   VAR 
      switching_on_inhibited : Bool := FALSE;
      ready_for_switching_on : Bool := FALSE;
      switched_on : Bool := FALSE;
      operation : Bool := FALSE;
      ars_statusword : Word;
      ars_controlword : Word;
      start_pos : Bool := FALSE;
      start_pos_old : Bool := FALSE;   // ***********************************************************************************************************************Anweisungsteil
      start_pos_man : Bool;
      start_pos_man_old : Bool;
      Fahrauftrag_OK : Bool;
      AFAG_Ist_Wert_in_Grad : Real;
      AFAG_soll_Wert_in_Grad : Real;
      AFAG_soll_Speed_in_Prozent : Int;
      AFAG_soll_Beschleunigung_in_Grad_s : Int;
      abs_rel : Bool;
      R_TRIG_Instance {InstructionName := 'R_TRIG'; LibVersion := '1.0'} : R_TRIG;
      R_TRIG_Q_Tipp_neg : Bool;
      R_TRIG_Instance_1 {InstructionName := 'R_TRIG'; LibVersion := '1.0'} : R_TRIG;
      R_TRIG_Instance_2 {InstructionName := 'R_TRIG'; LibVersion := '1.0'} : R_TRIG;
      TP_Time_Pos_0 {InstructionName := 'TP_TIME'; LibVersion := '1.0'} : TP_TIME;
      TP_Time_Pos_1 {InstructionName := 'TP_TIME'; LibVersion := '1.0'} : TP_TIME;
      TP_Time_Pos_2 {InstructionName := 'TP_TIME'; LibVersion := '1.0'} : TP_TIME;
      TP_Time_Pos_3 {InstructionName := 'TP_TIME'; LibVersion := '1.0'} : TP_TIME;
      TP_Time_Pos_4 {InstructionName := 'TP_TIME'; LibVersion := '1.0'} : TP_TIME;
      TP_Time_Pos_5 {InstructionName := 'TP_TIME'; LibVersion := '1.0'} : TP_TIME;
      TP_Time_Pos_6 {InstructionName := 'TP_TIME'; LibVersion := '1.0'} : TP_TIME;
      TP_Time_Pos_7 {InstructionName := 'TP_TIME'; LibVersion := '1.0'} : TP_TIME;
      TP_Time_Pos_8 {InstructionName := 'TP_TIME'; LibVersion := '1.0'} : TP_TIME;
      TP_Time_Pos_9 {InstructionName := 'TP_TIME'; LibVersion := '1.0'} : TP_TIME;
      TP_Time_Pos_10 {InstructionName := 'TP_TIME'; LibVersion := '1.0'} : TP_TIME;
      TP_Time_Pos_11 {InstructionName := 'TP_TIME'; LibVersion := '1.0'} : TP_TIME;
      TP_Time_Pos_12 {InstructionName := 'TP_TIME'; LibVersion := '1.0'} : TP_TIME;
      TP_Time_Pos_13 {InstructionName := 'TP_TIME'; LibVersion := '1.0'} : TP_TIME;
      TP_Time_Pos_14 {InstructionName := 'TP_TIME'; LibVersion := '1.0'} : TP_TIME;
      TP_Time_Pos_15 {InstructionName := 'TP_TIME'; LibVersion := '1.0'} : TP_TIME;
   END_VAR


BEGIN
	
	
	//Ausgänge zuweisen
	#A_UDT_Afag_soll_Werte.Telegrammkennung := 16#e0;
	#A_Afag_ist_wert_Grad := #AFAG_Ist_Wert_in_Grad;
	#AFAG_Ist_Wert_in_Grad := (DINT_TO_REAL(#E_UDT_Afag_ist_Werte.actual_position)); // / 1.000000e+003;
	#A_UDT_Afag_soll_Werte.Zielposition := REAL_TO_DINT(#AFAG_soll_Wert_in_Grad); // * 1.000000e+003);
	#A_UDT_Afag_soll_Werte.Fahrgeschwindigkeit := INT_TO_DINT(#AFAG_soll_Speed_in_Prozent * (#E_I_Max_Speed_Grad_s / 100));
	#A_UDT_Afag_soll_Werte.Beschleunigung := INT_TO_DINT(#AFAG_soll_Beschleunigung_in_Grad_s);
	#E_A_UDT_Afag_Positionen.A_Softw_ES_min_Grad := 0;
	#E_A_UDT_Afag_Positionen.A_Softw_ES_max_Grad := 360000;
	#E_A_UDT_Afag_Positionen.A_Max_Speed_Grad_s := #E_I_Max_Speed_Grad_s;
	#E_A_UDT_Afag_Positionen.A_Max_Beschleunigung_Grad_s := #E_I_Max_Beschleunigung_Grad_s;
	
	
	//************************************************************************************************
	
	//Lesen Statusword
	//Einlesen des Istzustands der Statemachine
	
	//    #DB_nr_actual_value_word:= INT_TO_WORD(#DB_nr_actual_value);
	//    #ars_statusword := PEEK_WORD (area := 16#84,
	//                                  dbNumber :=#DB_nr_actual_value_word,
	//                                  byteOffset := 2);
	#ars_statusword := #E_UDT_Afag_ist_Werte.PROFIDRIVE_Statusword;
	
	//Lesen Controlword
	//
	//  #DB_nr_position_word:=  INT_TO_WORD(#DB_nr_position);
	//  #ars_controlword := PEEK_WORD (area := 16#84,
	//                                  dbNumber :=#DB_nr_position_word,
	//                                  byteOffset := 2);
	
	// #ars_controlword := #A_UDT_Afag_soll_Werte.PROFIDRIVE_Controlword;
	
	//Steuern der Statemachine, S1 -> S2 -> S3 -> S4
	
	IF (#switching_on_inhibited                          //wenn state "switching_on_inhibited"
	    AND #E_drive_enable)                             //und  Reglerfreigabe
	THEN
	    #ars_controlword := 16#0406;              //dann state "ready_for_switching_on" anfordern,
	ELSIF (#switching_on_inhibited                     //
	    AND (NOT (#E_drive_enable)))                      //wenn Reglerfreigabe aus,
	THEN
	    #ars_controlword := 16#0400;              //dann state "switching_on_inhibited" anfordern.
	END_IF;
	
	IF (#ready_for_switching_on                          //wenn state "ready_for_switching_on"
	    AND #E_drive_enable)                             //und Reglerfeigabe
	THEN
	    #ars_controlword := 16#0407;              //dann state "switched_on" anfordern,
	ELSIF (#ready_for_switching_on                     //
	    AND (NOT (#E_drive_enable)))                      //wenn Reglerfeigabe aus,
	THEN
	    #ars_controlword := 16#0400;              //dann state "switching_on_inhibited" anfordern.
	END_IF;
	
	IF (#switched_on                                     //wenn state "switched_on"
	    AND #E_drive_enable)                             //und Reglerfeigabe
	THEN
	    #ars_controlword := 16#040f;              //dann state "operation" anfordern,
	ELSIF (#switched_on                                //
	    AND (NOT (#E_drive_enable)))                      //wenn Reglerfeigabe aus,
	THEN
	    #ars_controlword := 16#0400;              //dann state "switching_on_inhibited" anfordern.
	END_IF;
	
	IF (#operation                                       //wenn state "operation"
	    AND (NOT (#E_drive_enable)))                      //und keine Reglerfeigabe
	THEN
	    #ars_controlword := 16#040e;              //dann state "switching_on_inhibited" anfordern.
	END_IF;
	
	//************************************************************************************************
	
	//Kommandos über digitale Eingänge
	// Bit 10 (control by plc) im Controlword muss immer gesetzt sein
	
	IF #E_start_homing
	THEN
	    #ars_controlword := (#ars_controlword OR 16#0C00);    //Setzen Bit 11 im STW1
	ELSE
	    #ars_controlword := (#ars_controlword & 16#f7ff);
	END_IF;
	
	IF (#Fahrauftrag_OK = 1) THEN
	    IF (#start_pos_old <> #start_pos) OR (#start_pos_man_old <> #start_pos_man)
	    THEN
	        IF #start_pos OR #start_pos_man
	        THEN
	            #ars_controlword := (#ars_controlword OR 16#0440);    //Setzen Bit 6 im STW1
	        ELSE
	            #ars_controlword := (#ars_controlword & 16#ffbf);
	        END_IF;
	    END_IF;
	    
	    #start_pos_old := #start_pos;
	    #start_pos_man_old := #start_pos_man;
	    
	END_IF;
	
	
	
	
	IF #abs_rel
	THEN
	    #ars_controlword := (#ars_controlword OR 16#1400);   //Setzen Bit 12 im STW1
	ELSE
	    #ars_controlword := (#ars_controlword & 16#efff);
	END_IF;
	
	IF #E_change_immediatly
	THEN
	    #ars_controlword := (#ars_controlword OR 16#2400);   //Setzen Bit 13 im STW1
	ELSE
	    #ars_controlword := (#ars_controlword & 16#dfff);
	END_IF;
	
	IF #E_intermediate_stop
	THEN
	    #ars_controlword := (#ars_controlword & 16#ffdf);   //Rücksetzen Bit 5 im STW1
	ELSE
	    #ars_controlword := (#ars_controlword OR 16#0420);
	END_IF;
	
	IF #E_hold
	THEN
	    #ars_controlword := (#ars_controlword & 16#ffef);    //Rücksetzen Bit 4 im STW1
	    #ars_controlword := (#ars_controlword & 16#feff);    //Rücksetzen jog_pos
	    #ars_controlword := (#ars_controlword & 16#fdff);    //Rücksetzen jog_neg
	ELSE
	    #ars_controlword := (#ars_controlword OR 16#0410);
	END_IF;
	
	IF (#E_jog_pos AND NOT #E_hold)
	THEN
	    #ars_controlword := (#ars_controlword OR 16#0500);    //Setzen Bit 8 im STW1
	ELSE
	    #ars_controlword := (#ars_controlword & 16#feff);
	END_IF;
	
	IF (#E_jog_neg AND NOT #E_hold)
	THEN
	    #ars_controlword := (#ars_controlword OR 16#0600);    //Setzen Bit 9 im STW1
	ELSE
	    #ars_controlword := (#ars_controlword & 16#fdff);
	END_IF;
	
	IF #E_fault_reset
	THEN
	    #ars_controlword := (#ars_controlword OR 16#0480);    //Setzen Bit 7 im STW1
	ELSE
	    #ars_controlword := (#ars_controlword & 16#ff7f);
	END_IF;
	
	
	//************************************************************************************************
	
	//Setzen digitaler Ausgänge
	
	IF #operation
	THEN
	    #A_drive_enable_ok := TRUE;
	ELSE
	    #A_drive_enable_ok := FALSE;
	END_IF;
	
	IF ((#ars_statusword & 16#0800) = 16#0800)    //Bit 11 vom ZSW1
	THEN
	    #A_home_valid := TRUE;
	ELSE
	    #A_home_valid := FALSE;
	END_IF;
	
	IF ((#ars_statusword & 16#0400) = 16#0400)    //Bit 10 vom ZSW1
	THEN
	    #A_pos_ok := TRUE;
	ELSE
	    #A_pos_ok := FALSE;
	END_IF;
	
	IF ((#ars_statusword & 16#2000) = 16#2000)    //Bit 13 vom ZSW1
	THEN
	    #A_velo_zero := TRUE;
	ELSE
	    #A_velo_zero := FALSE;
	END_IF;
	
	IF ((#ars_statusword & 16#0008) = 16#0008)    //Bit 3 vom ZSW1
	THEN
	    #A_fault := TRUE;
	ELSE
	    #A_fault := FALSE;
	END_IF;
	
	//************************************************************************************************
	
	//Schreiben Controlword
	
	//  POKE (area := 16#84,
	//        dbNumber := #DB_nr_position_word,
	//        byteOffset := 2,
	//        value := #ars_controlword );
	
	#A_UDT_Afag_soll_Werte.PROFIDRIVE_Controlword := #ars_controlword;
	
	
	// Achse mit Position Starten
	// Position[0]
	
	    IF #E_A_UDT_Afag_Positionen.Start_POS_Position[0] THEN
	    #AFAG_soll_Wert_in_Grad := #E_A_UDT_Afag_Positionen.Soll_Wert_in_Grad_Position[0];
	    #AFAG_soll_Beschleunigung_in_Grad_s := #E_A_UDT_Afag_Positionen.Soll_Beschleunigung_in_Grad_s_Position[0];
	    #start_pos := true;
	    
	    #AFAG_soll_Speed_in_Prozent := #E_A_UDT_Afag_Positionen.Soll_Speed_in_Prozent_Position[0];
	END_IF;
	
	// Position[1]
	
	IF #E_A_UDT_Afag_Positionen.Start_POS_Position[1] THEN
	    #AFAG_soll_Wert_in_Grad := #E_A_UDT_Afag_Positionen.Soll_Wert_in_Grad_Position[1];
	    #AFAG_soll_Beschleunigung_in_Grad_s := #E_A_UDT_Afag_Positionen.Soll_Beschleunigung_in_Grad_s_Position[1];
	    #start_pos := true;
	    
	    #AFAG_soll_Speed_in_Prozent := #E_A_UDT_Afag_Positionen.Soll_Speed_in_Prozent_Position[1];
	END_IF;
	
	
	// Position 2
	
	IF #E_A_UDT_Afag_Positionen.Start_POS_Position[2] THEN
	    #AFAG_soll_Wert_in_Grad := #E_A_UDT_Afag_Positionen.Soll_Wert_in_Grad_Position[2];
	    #AFAG_soll_Beschleunigung_in_Grad_s := #E_A_UDT_Afag_Positionen.Soll_Beschleunigung_in_Grad_s_Position[2];
	    #start_pos := true;
	    
	    #AFAG_soll_Speed_in_Prozent := #E_A_UDT_Afag_Positionen.Soll_Speed_in_Prozent_Position[2];
	END_IF;
	
	// Position 3
	
	IF #E_A_UDT_Afag_Positionen.Start_POS_Position[3] THEN
	    #AFAG_soll_Wert_in_Grad := #E_A_UDT_Afag_Positionen.Soll_Wert_in_Grad_Position[3];
	    #AFAG_soll_Beschleunigung_in_Grad_s := #E_A_UDT_Afag_Positionen.Soll_Beschleunigung_in_Grad_s_Position[3];
	    #start_pos := true;
	    
	    #AFAG_soll_Speed_in_Prozent := #E_A_UDT_Afag_Positionen.Soll_Speed_in_Prozent_Position[3];
	END_IF;
	
	// Position 4
	
	IF #E_A_UDT_Afag_Positionen.Start_POS_Position[4] THEN
	    #AFAG_soll_Wert_in_Grad := #E_A_UDT_Afag_Positionen.Soll_Wert_in_Grad_Position[4];
	    #AFAG_soll_Beschleunigung_in_Grad_s := #E_A_UDT_Afag_Positionen.Soll_Beschleunigung_in_Grad_s_Position[4];
	    #start_pos := true;
	    
	    #AFAG_soll_Speed_in_Prozent := #E_A_UDT_Afag_Positionen.Soll_Speed_in_Prozent_Position[4];
	END_IF;
	
	// Position 5
	
	IF #E_A_UDT_Afag_Positionen.Start_POS_Position[5] THEN
	    #AFAG_soll_Wert_in_Grad := #E_A_UDT_Afag_Positionen.Soll_Wert_in_Grad_Position[5];
	    #AFAG_soll_Beschleunigung_in_Grad_s := #E_A_UDT_Afag_Positionen.Soll_Beschleunigung_in_Grad_s_Position[5];
	    #start_pos := true;
	    
	    #AFAG_soll_Speed_in_Prozent := #E_A_UDT_Afag_Positionen.Soll_Speed_in_Prozent_Position[5];
	END_IF;
	
	// Position 6
	
	IF #E_A_UDT_Afag_Positionen.Start_POS_Position[6] THEN
	    #AFAG_soll_Wert_in_Grad := #E_A_UDT_Afag_Positionen.Soll_Wert_in_Grad_Position[6];
	    #AFAG_soll_Beschleunigung_in_Grad_s := #E_A_UDT_Afag_Positionen.Soll_Beschleunigung_in_Grad_s_Position[6];
	    #start_pos := true;
	    
	    #AFAG_soll_Speed_in_Prozent := #E_A_UDT_Afag_Positionen.Soll_Speed_in_Prozent_Position[6];
	END_IF;
	
	// Position 7
	
	IF #E_A_UDT_Afag_Positionen.Start_POS_Position[7] THEN
	    #AFAG_soll_Wert_in_Grad := #E_A_UDT_Afag_Positionen.Soll_Wert_in_Grad_Position[7];
	    #AFAG_soll_Beschleunigung_in_Grad_s := #E_A_UDT_Afag_Positionen.Soll_Beschleunigung_in_Grad_s_Position[7];
	    #start_pos := true;
	    
	    #AFAG_soll_Speed_in_Prozent := #E_A_UDT_Afag_Positionen.Soll_Speed_in_Prozent_Position[7];
	END_IF;
	
	// Position 8
	
	IF #E_A_UDT_Afag_Positionen.Start_POS_Position[8] THEN
	    #AFAG_soll_Wert_in_Grad := #E_A_UDT_Afag_Positionen.Soll_Wert_in_Grad_Position[8];
	    #AFAG_soll_Beschleunigung_in_Grad_s := #E_A_UDT_Afag_Positionen.Soll_Beschleunigung_in_Grad_s_Position[8];
	    #start_pos := true;
	    
	    #AFAG_soll_Speed_in_Prozent := #E_A_UDT_Afag_Positionen.Soll_Speed_in_Prozent_Position[8];
	END_IF;
	
	// Position 9
	
	IF #E_A_UDT_Afag_Positionen.Start_POS_Position[9] THEN
	    #AFAG_soll_Wert_in_Grad := #E_A_UDT_Afag_Positionen.Soll_Wert_in_Grad_Position[9];
	    #AFAG_soll_Beschleunigung_in_Grad_s := #E_A_UDT_Afag_Positionen.Soll_Beschleunigung_in_Grad_s_Position[9];
	    #start_pos := true;
	   
	    #AFAG_soll_Speed_in_Prozent := #E_A_UDT_Afag_Positionen.Soll_Speed_in_Prozent_Position[9];
	END_IF;
	
	// Position 10
	
	IF #E_A_UDT_Afag_Positionen.Start_POS_Position[10] THEN
	    #AFAG_soll_Wert_in_Grad := #E_A_UDT_Afag_Positionen.Soll_Wert_in_Grad_Position[10];
	    #AFAG_soll_Beschleunigung_in_Grad_s := #E_A_UDT_Afag_Positionen.Soll_Beschleunigung_in_Grad_s_Position[10];
	    #start_pos := true;
	    
	    #AFAG_soll_Speed_in_Prozent := #E_A_UDT_Afag_Positionen.Soll_Speed_in_Prozent_Position[10];
	END_IF;
	
	// Position 11
	
	IF #E_A_UDT_Afag_Positionen.Start_POS_Position[11] THEN
	    #AFAG_soll_Wert_in_Grad := #E_A_UDT_Afag_Positionen.Soll_Wert_in_Grad_Position[11];
	    #AFAG_soll_Beschleunigung_in_Grad_s := #E_A_UDT_Afag_Positionen.Soll_Beschleunigung_in_Grad_s_Position[11];
	    #start_pos := true;
	    
	    #AFAG_soll_Speed_in_Prozent := #E_A_UDT_Afag_Positionen.Soll_Speed_in_Prozent_Position[11];
	END_IF;
	
	// Position 12
	
	IF #E_A_UDT_Afag_Positionen.Start_POS_Position[12] THEN
	    #AFAG_soll_Wert_in_Grad := #E_A_UDT_Afag_Positionen.Soll_Wert_in_Grad_Position[12];
	    #AFAG_soll_Beschleunigung_in_Grad_s := #E_A_UDT_Afag_Positionen.Soll_Beschleunigung_in_Grad_s_Position[12];
	    #start_pos := true;
	    
	    #AFAG_soll_Speed_in_Prozent := #E_A_UDT_Afag_Positionen.Soll_Speed_in_Prozent_Position[12];
	END_IF;
	
	// Position 13
	
	IF #E_A_UDT_Afag_Positionen.Start_POS_Position[13] THEN
	    #AFAG_soll_Wert_in_Grad := #E_A_UDT_Afag_Positionen.Soll_Wert_in_Grad_Position[13];
	    #AFAG_soll_Beschleunigung_in_Grad_s := #E_A_UDT_Afag_Positionen.Soll_Beschleunigung_in_Grad_s_Position[13];
	    #start_pos := true;
	    
	    #AFAG_soll_Speed_in_Prozent := #E_A_UDT_Afag_Positionen.Soll_Speed_in_Prozent_Position[13];
	END_IF;
	
	// Position 14
	
	IF #E_A_UDT_Afag_Positionen.Start_POS_Position[14] THEN
	    #AFAG_soll_Wert_in_Grad := #E_A_UDT_Afag_Positionen.Soll_Wert_in_Grad_Position[14];
	    #AFAG_soll_Beschleunigung_in_Grad_s := #E_A_UDT_Afag_Positionen.Soll_Beschleunigung_in_Grad_s_Position[14];
	    #start_pos := true;
	    
	    #AFAG_soll_Speed_in_Prozent := #E_A_UDT_Afag_Positionen.Soll_Speed_in_Prozent_Position[14];
	END_IF;
	
	// Position 15
	
	IF #E_A_UDT_Afag_Positionen.Start_POS_Position[15] THEN
	    #AFAG_soll_Wert_in_Grad := #E_A_UDT_Afag_Positionen.Soll_Wert_in_Grad_Position[15];
	    #AFAG_soll_Beschleunigung_in_Grad_s := #E_A_UDT_Afag_Positionen.Soll_Beschleunigung_in_Grad_s_Position[15];
	    #start_pos := true;
	    
	    #AFAG_soll_Speed_in_Prozent := #E_A_UDT_Afag_Positionen.Soll_Speed_in_Prozent_Position[15];
	END_IF;
	
	// Manuelle Geschwindigkeitsanpassung
	IF #E_BA_Manuell = TRUE THEN
	   #AFAG_soll_Speed_in_Prozent := #E_I_Manuell_Geschwindigkeit_Prozent;
	   #AFAG_soll_Beschleunigung_in_Grad_s := 1000;
	END_IF;
	
	IF( (#E_A_UDT_Afag_Positionen.Start_POS_Position[0] AND #E_A_UDT_Afag_Positionen.POS_OK_Position[0])OR
	   (#E_A_UDT_Afag_Positionen.Start_POS_Position[1]AND #E_A_UDT_Afag_Positionen.POS_OK_Position[1])OR
	   (#E_A_UDT_Afag_Positionen.Start_POS_Position[2]AND #E_A_UDT_Afag_Positionen.POS_OK_Position[2])OR
	   (#E_A_UDT_Afag_Positionen.Start_POS_Position[3]AND #E_A_UDT_Afag_Positionen.POS_OK_Position[3])OR
	   (#E_A_UDT_Afag_Positionen.Start_POS_Position[4]AND #E_A_UDT_Afag_Positionen.POS_OK_Position[4])OR
	   (#E_A_UDT_Afag_Positionen.Start_POS_Position[5]AND #E_A_UDT_Afag_Positionen.POS_OK_Position[5])OR
	   (#E_A_UDT_Afag_Positionen.Start_POS_Position[6]AND #E_A_UDT_Afag_Positionen.POS_OK_Position[6])OR
	   (#E_A_UDT_Afag_Positionen.Start_POS_Position[7]AND #E_A_UDT_Afag_Positionen.POS_OK_Position[7])OR
	   (#E_A_UDT_Afag_Positionen.Start_POS_Position[8]AND #E_A_UDT_Afag_Positionen.POS_OK_Position[8])OR
	   (#E_A_UDT_Afag_Positionen.Start_POS_Position[9]AND #E_A_UDT_Afag_Positionen.POS_OK_Position[9])OR
	   (#E_A_UDT_Afag_Positionen.Start_POS_Position[10]AND #E_A_UDT_Afag_Positionen.POS_OK_Position[10])OR
	   (#E_A_UDT_Afag_Positionen.Start_POS_Position[11]AND #E_A_UDT_Afag_Positionen.POS_OK_Position[11])OR
	   (#E_A_UDT_Afag_Positionen.Start_POS_Position[12]AND #E_A_UDT_Afag_Positionen.POS_OK_Position[12])OR
	   (#E_A_UDT_Afag_Positionen.Start_POS_Position[13]AND #E_A_UDT_Afag_Positionen.POS_OK_Position[13])OR
	   (#E_A_UDT_Afag_Positionen.Start_POS_Position[14]AND #E_A_UDT_Afag_Positionen.POS_OK_Position[14])OR
	   (#E_A_UDT_Afag_Positionen.Start_POS_Position[15]AND #E_A_UDT_Afag_Positionen.POS_OK_Position[15])OR
	    #E_Richten_reset_FRG)
	THEN
	    #start_pos := 0;
	    #E_A_UDT_Afag_Positionen.Start_POS_Position[0] := 0;
	    #E_A_UDT_Afag_Positionen.Start_POS_Position[1] := 0;
	    #E_A_UDT_Afag_Positionen.Start_POS_Position[2] := 0;
	    #E_A_UDT_Afag_Positionen.Start_POS_Position[3] := 0;
	    #E_A_UDT_Afag_Positionen.Start_POS_Position[4] := 0;
	    #E_A_UDT_Afag_Positionen.Start_POS_Position[5] := 0;
	    #E_A_UDT_Afag_Positionen.Start_POS_Position[6] := 0;
	    #E_A_UDT_Afag_Positionen.Start_POS_Position[7] := 0;
	    #E_A_UDT_Afag_Positionen.Start_POS_Position[8] := 0;
	    #E_A_UDT_Afag_Positionen.Start_POS_Position[9] := 0;
	    #E_A_UDT_Afag_Positionen.Start_POS_Position[10] := 0;
	    #E_A_UDT_Afag_Positionen.Start_POS_Position[11] := 0;
	    #E_A_UDT_Afag_Positionen.Start_POS_Position[12] := 0;
	    #E_A_UDT_Afag_Positionen.Start_POS_Position[13] := 0;
	    #E_A_UDT_Afag_Positionen.Start_POS_Position[14] := 0;
	    #E_A_UDT_Afag_Positionen.Start_POS_Position[15] := 0;
	    #E_A_UDT_Afag_Positionen.POS_OK_Position[15] := 0;
	END_IF;
	
	
	// Achse Positionsrückmeldung
	
	IF #E_A_UDT_Afag_Positionen.Start_POS_Position[0] AND #A_pos_ok
	THEN
	    #E_A_UDT_Afag_Positionen.POS_OK_Position[0] := 1;
	ELSE
	    #E_A_UDT_Afag_Positionen.POS_OK_Position[0] := 0;
	END_IF;
	
	IF #E_A_UDT_Afag_Positionen.Start_POS_Position[1] AND #A_pos_ok
	THEN
	    #E_A_UDT_Afag_Positionen.POS_OK_Position[1] := 1;
	ELSE
	    #E_A_UDT_Afag_Positionen.POS_OK_Position[1] := 0;
	END_IF;
	
	IF #E_A_UDT_Afag_Positionen.Start_POS_Position[2] AND #A_pos_ok
	THEN
	    #E_A_UDT_Afag_Positionen.POS_OK_Position[2] := 1;
	ELSE
	    #E_A_UDT_Afag_Positionen.POS_OK_Position[2] := 0;
	END_IF;
	
	IF #E_A_UDT_Afag_Positionen.Start_POS_Position[3] AND #A_pos_ok
	THEN
	    #E_A_UDT_Afag_Positionen.POS_OK_Position[3] := 1;
	ELSE
	    #E_A_UDT_Afag_Positionen.POS_OK_Position[3] := 0;
	END_IF;
	
	IF #E_A_UDT_Afag_Positionen.Start_POS_Position[4] AND #A_pos_ok
	THEN
	    #E_A_UDT_Afag_Positionen.POS_OK_Position[4] := 1;
	ELSE
	    #E_A_UDT_Afag_Positionen.POS_OK_Position[4] := 0;
	END_IF;
	
	IF #E_A_UDT_Afag_Positionen.Start_POS_Position[5] AND #A_pos_ok
	THEN
	    #E_A_UDT_Afag_Positionen.POS_OK_Position[5] := 1;
	ELSE
	    #E_A_UDT_Afag_Positionen.POS_OK_Position[5] := 0;
	END_IF;
	
	IF #E_A_UDT_Afag_Positionen.Start_POS_Position[6] AND #A_pos_ok
	THEN
	    #E_A_UDT_Afag_Positionen.POS_OK_Position[6] := 1;
	ELSE
	    #E_A_UDT_Afag_Positionen.POS_OK_Position[6] := 0;
	END_IF;
	
	IF #E_A_UDT_Afag_Positionen.Start_POS_Position[7] AND #A_pos_ok
	THEN
	    #E_A_UDT_Afag_Positionen.POS_OK_Position[7] := 1;
	ELSE
	    #E_A_UDT_Afag_Positionen.POS_OK_Position[7] := 0;
	END_IF;
	
	IF #E_A_UDT_Afag_Positionen.Start_POS_Position[8] AND #A_pos_ok
	THEN
	    #E_A_UDT_Afag_Positionen.POS_OK_Position[8] := 1;
	ELSE
	    #E_A_UDT_Afag_Positionen.POS_OK_Position[8] := 0;
	END_IF;
	
	IF #E_A_UDT_Afag_Positionen.Start_POS_Position[9] AND #A_pos_ok
	THEN
	    #E_A_UDT_Afag_Positionen.POS_OK_Position[9] := 1;
	ELSE
	    #E_A_UDT_Afag_Positionen.POS_OK_Position[9] := 0;
	END_IF;
	
	IF #E_A_UDT_Afag_Positionen.Start_POS_Position[10] AND #A_pos_ok
	THEN
	    #E_A_UDT_Afag_Positionen.POS_OK_Position[10] := 1;
	ELSE
	    #E_A_UDT_Afag_Positionen.POS_OK_Position[10] := 0;
	END_IF;
	
	IF #E_A_UDT_Afag_Positionen.Start_POS_Position[11] AND #A_pos_ok
	THEN
	    #E_A_UDT_Afag_Positionen.POS_OK_Position[11] := 1;
	ELSE
	    #E_A_UDT_Afag_Positionen.POS_OK_Position[11] := 0;
	END_IF;
	
	IF #E_A_UDT_Afag_Positionen.Start_POS_Position[12] AND #A_pos_ok
	THEN
	    #E_A_UDT_Afag_Positionen.POS_OK_Position[12] := 1;
	ELSE
	    #E_A_UDT_Afag_Positionen.POS_OK_Position[12] := 0;
	END_IF;
	
	IF #E_A_UDT_Afag_Positionen.Start_POS_Position[13] AND #A_pos_ok
	THEN
	    #E_A_UDT_Afag_Positionen.POS_OK_Position[13] := 1;
	ELSE
	    #E_A_UDT_Afag_Positionen.POS_OK_Position[13] := 0;
	END_IF;
	
	IF #E_A_UDT_Afag_Positionen.Start_POS_Position[14] AND #A_pos_ok
	THEN
	    #E_A_UDT_Afag_Positionen.POS_OK_Position[14] := 1;
	ELSE
	    #E_A_UDT_Afag_Positionen.POS_OK_Position[14] := 0;
	END_IF;
	
	IF #E_A_UDT_Afag_Positionen.Start_POS_Position[15] AND #A_pos_ok
	THEN
	    #E_A_UDT_Afag_Positionen.POS_OK_Position[15] := 1;
	ELSE
	    #E_A_UDT_Afag_Positionen.POS_OK_Position[15] := 0;
	END_IF;
	
	IF
	    (#E_A_UDT_Afag_Positionen.Start_POS_Position[0]) OR
	    (#E_A_UDT_Afag_Positionen.Start_POS_Position[1]) OR
	    (#E_A_UDT_Afag_Positionen.Start_POS_Position[2]) OR
	    (#E_A_UDT_Afag_Positionen.Start_POS_Position[3]) OR
	    (#E_A_UDT_Afag_Positionen.Start_POS_Position[4]) OR
	    (#E_A_UDT_Afag_Positionen.Start_POS_Position[5]) OR
	    (#E_A_UDT_Afag_Positionen.Start_POS_Position[6]) OR
	    (#E_A_UDT_Afag_Positionen.Start_POS_Position[7]) OR
	    (#E_A_UDT_Afag_Positionen.Start_POS_Position[8]) OR
	    (#E_A_UDT_Afag_Positionen.Start_POS_Position[9]) OR
	    (#E_A_UDT_Afag_Positionen.Start_POS_Position[10]) OR
	    (#E_A_UDT_Afag_Positionen.Start_POS_Position[11]) OR
	    (#E_A_UDT_Afag_Positionen.Start_POS_Position[12]) OR
	    (#E_A_UDT_Afag_Positionen.Start_POS_Position[13]) OR
	    (#E_A_UDT_Afag_Positionen.Start_POS_Position[14]) OR
	    (#E_A_UDT_Afag_Positionen.Start_POS_Position[15]) OR
	    (#start_pos)
	THEN
	    #A_Fahrauftrag_Aktiv := 1;
	ELSE
	    #A_Fahrauftrag_Aktiv := 0;
	END_IF;
	
	
	
	
	//Reset Start pos
	IF ((#A_pos_ok = true) OR (#A_drive_enable_ok = FALSE) OR (#E_fault_reset = TRUE))
	THEN
	    #start_pos_man := false;
	    #abs_rel := true;
	END_IF;
	
	//Tipp pos
	#R_TRIG_Instance(CLK:=#E_Tipp_pos);
	IF (#R_TRIG_Instance.Q AND NOT #start_pos_man)
	THEN
	    #AFAG_soll_Wert_in_Grad := #E_R_Verfahrweg_Grad;
	    #start_pos_man := TRUE;
	END_IF;
	
	//Tipp neg
	#R_TRIG_Instance_1(CLK:=#E_Tipp_neg);
	IF (#R_TRIG_Instance_1.Q AND NOT #start_pos_man)
	THEN
	    #AFAG_soll_Wert_in_Grad := #E_R_Verfahrweg_Grad;
	    #start_pos_man := TRUE;
	END_IF;
	
	//absolut verfahren
	#R_TRIG_Instance_2(CLK:=#E_Start_pos_man);
	IF(#R_TRIG_Instance_2.Q AND NOT #start_pos_man)
	THEN
	    #AFAG_soll_Wert_in_Grad := #E_R_Afag_soll_wert_man_Grad;
	    #start_pos_man := TRUE;
	    #abs_rel := false;
	END_IF;
	
	// keine Endlagenüberwachung bei Drehachse
	// Überwachung Fahrauftrag
	    #Fahrauftrag_OK := TRUE;
	 
	    
	//Einlesen des Istzustands der Statemachine
	   IF ((#ars_statusword & 16#0047) = 16#0040)
	        THEN #switching_on_inhibited := TRUE;
	        ELSE #switching_on_inhibited := FALSE;
	    END_IF;
	
	    IF ((#ars_statusword & 16#0047) = 16#0001)
	        THEN #ready_for_switching_on:= TRUE;
	        ELSE #ready_for_switching_on:= FALSE;
	    END_IF;
	     
	    IF ((#ars_statusword & 16#0047) = 16#0003)
	        THEN #switched_on:= TRUE;
	        ELSE #switched_on:= FALSE;
	    END_IF;
	
	    IF ((#ars_statusword & 16#0047) = 16#0007)
	        THEN #operation:= TRUE;
	        ELSE #operation:= FALSE;
	    END_IF;    
	
	
	
	    
	    
END_FUNCTION_BLOCK

FUNCTION_BLOCK "BB_Ansteuerung_Afag_offen_V02.3"
TITLE = 'FB Positionierbetrieb'
{ S7_Optimized_Access := 'TRUE' }
AUTHOR : Essmann
FAMILY : metronix
NAME : position
VERSION : 1.1
//Der Baustein kann nicht rückübersetzt und unter STEP7 bearbeitet werden.  Der Baustein kann nur als Quelle im Ordner "Quellen" bearbeitet werden.    IO-Variablen  
   VAR_INPUT 
      drive_enable : Bool := FALSE;
      start_homing : Bool := FALSE;
      start_pos : Bool := FALSE;
      abs_rel : Bool := FALSE;
      change_immediatly : Bool := FALSE;
      intermediate_stop : Bool := FALSE;
      hold : Bool := FALSE;
      jog_pos : Bool := FALSE;
      jog_neg : Bool := FALSE;
      fault_reset : Bool := FALSE;
      E_Afag_ist_Werte : "Afag_ist_Werte";
   END_VAR

   VAR_OUTPUT 
      drive_enable_ok : Bool := FALSE;
      home_valid : Bool := FALSE;
      pos_ok : Bool := FALSE;
      velo_zero : Bool := FALSE;
      fault : Bool := FALSE;   // statische Variablen
   END_VAR

   VAR_IN_OUT 
      A_Afag_soll_Werte : "Afag_soll_Werte";
   END_VAR

   VAR 
      DB_nr_position_word : Word;
      DB_nr_actual_value_word : Word;
      switching_on_inhibited : Bool := FALSE;
      ready_for_switching_on : Bool := FALSE;
      switched_on : Bool := FALSE;
      operation : Bool := FALSE;
      ars_statusword : Word;
      ars_controlword : Word;
      start_pos_old : Bool := FALSE;   // ***********************************************************************************************************************Anweisungsteil
   END_VAR


BEGIN
	
	
	//Lesen Statusword
	//Einlesen des Istzustands der Statemachine
	    
	 //    #DB_nr_actual_value_word:= INT_TO_WORD(#DB_nr_actual_value);
	 //    #ars_statusword := PEEK_WORD (area := 16#84,
	 //                                  dbNumber :=#DB_nr_actual_value_word,
	 //                                  byteOffset := 2);
	 
	 #A_Afag_soll_Werte.Telegrammkennung:= 16#e0;
	 
	 
	 #ars_statusword := #E_Afag_ist_Werte.PROFIDRIVE_Statusword;
	
	   IF ((#ars_statusword & 16#0047) = 16#0040)
	        THEN #switching_on_inhibited := TRUE;
	        ELSE #switching_on_inhibited := FALSE;
	    END_IF;
	
	    IF ((#ars_statusword & 16#0047) = 16#0001)
	        THEN #ready_for_switching_on:= TRUE;
	        ELSE #ready_for_switching_on:= FALSE;
	    END_IF;
	     
	    IF ((#ars_statusword & 16#0047) = 16#0003)
	        THEN #switched_on:= TRUE;
	        ELSE #switched_on:= FALSE;
	    END_IF;
	
	    IF ((#ars_statusword & 16#0047) = 16#0007)
	        THEN #operation:= TRUE;
	        ELSE #operation:= FALSE;
	    END_IF;    
	
	
	//************************************************************************************************
	
	//Lesen Controlword
	//
	 //  #DB_nr_position_word:=  INT_TO_WORD(#DB_nr_position);
	 //  #ars_controlword := PEEK_WORD (area := 16#84,
	 //                                  dbNumber :=#DB_nr_position_word,
	 //                                  byteOffset := 2);
	    
	    #ars_controlword := #A_Afag_soll_Werte.PROFIDRIVE_Controlword;
	    
	//Steuern der Statemachine, S1 -> S2 -> S3 -> S4
	
	  IF (#switching_on_inhibited                          //wenn state "switching_on_inhibited"
	        AND #drive_enable)                             //und  Reglerfreigabe
	        THEN #ars_controlword := 16#0406;              //dann state "ready_for_switching_on" anfordern,
	    ELSIF (#switching_on_inhibited                     //
	        AND (NOT(#drive_enable)))                      //wenn Reglerfreigabe aus,
	        THEN #ars_controlword := 16#0400;              //dann state "switching_on_inhibited" anfordern.
	  END_IF;                                             
	
	  IF (#ready_for_switching_on                          //wenn state "ready_for_switching_on"
	        AND #drive_enable)                             //und Reglerfeigabe
	        THEN #ars_controlword := 16#0407;              //dann state "switched_on" anfordern,
	    ELSIF (#ready_for_switching_on                     //
	        AND (NOT(#drive_enable)))                      //wenn Reglerfeigabe aus,
	        THEN #ars_controlword := 16#0400;              //dann state "switching_on_inhibited" anfordern.
	  END_IF;
	
	  IF (#switched_on                                     //wenn state "switched_on"
	        AND #drive_enable)                             //und Reglerfeigabe
	        THEN #ars_controlword := 16#040f;              //dann state "operation" anfordern,
	    ELSIF (#switched_on                                //
	        AND (NOT(#drive_enable)))                      //wenn Reglerfeigabe aus,
	        THEN #ars_controlword := 16#0400;              //dann state "switching_on_inhibited" anfordern.
	  END_IF;
	
	  IF (#operation                                       //wenn state "operation"
	        AND (NOT(#drive_enable)))                      //und keine Reglerfeigabe
	        THEN #ars_controlword := 16#040e;              //dann state "switching_on_inhibited" anfordern.
	  END_IF;
	
	//************************************************************************************************
	
	//Kommandos über digitale Eingänge
	// Bit 10 (control by plc) im Controlword muss immer gesetzt sein
	
	    IF #start_homing
	        THEN #ars_controlword := (#ars_controlword OR 16#0C00);    //Setzen Bit 11 im STW1
	        ELSE #ars_controlword := (#ars_controlword  & 16#f7ff);
	    END_IF;
	
	    IF #start_pos_old <> #start_pos
	        THEN IF #start_pos 
	                 THEN #ars_controlword := (#ars_controlword OR 16#0440);    //Setzen Bit 6 im STW1
	                 ELSE #ars_controlword := (#ars_controlword  & 16#ffbf);
	             END_IF;
	    END_IF;
	
	    #start_pos_old := #start_pos;
	
	    IF #abs_rel
	        THEN #ars_controlword := (#ars_controlword OR 16#1400);   //Setzen Bit 12 im STW1
	        ELSE #ars_controlword := (#ars_controlword  & 16#efff);
	    END_IF;
	    
	    IF #change_immediatly
	        THEN #ars_controlword := (#ars_controlword OR 16#2400);   //Setzen Bit 13 im STW1
	        ELSE #ars_controlword := (#ars_controlword  & 16#dfff);
	    END_IF;
	   
	    IF #intermediate_stop
	        THEN #ars_controlword := (#ars_controlword  & 16#ffdf);   //Rücksetzen Bit 5 im STW1
	        ELSE #ars_controlword := (#ars_controlword OR 16#0420);
	    END_IF;
	
	    IF #hold
	        THEN #ars_controlword := (#ars_controlword  & 16#ffef);    //Rücksetzen Bit 4 im STW1
	             #ars_controlword := (#ars_controlword  & 16#feff);    //Rücksetzen jog_pos
	             #ars_controlword := (#ars_controlword  & 16#fdff);    //Rücksetzen jog_neg
	        ELSE #ars_controlword := (#ars_controlword OR 16#0410);
	    END_IF;
	
	    IF (#jog_pos AND NOT #hold)
	        THEN #ars_controlword := (#ars_controlword OR 16#0500);    //Setzen Bit 8 im STW1
	        ELSE #ars_controlword := (#ars_controlword  & 16#feff);
	    END_IF;
	
	    IF (#jog_neg AND NOT #hold)
	        THEN #ars_controlword := (#ars_controlword OR 16#0600);    //Setzen Bit 9 im STW1
	        ELSE #ars_controlword := (#ars_controlword  & 16#fdff);
	    END_IF;
	
	    IF #fault_reset
	        THEN #ars_controlword := (#ars_controlword OR 16#0480);    //Setzen Bit 7 im STW1
	        ELSE #ars_controlword := (#ars_controlword  & 16#ff7f);
	    END_IF;
	
	
	//************************************************************************************************
	
	//Setzen digitaler Ausgänge
	
	    IF #operation
	        THEN #drive_enable_ok := TRUE;
	        ELSE #drive_enable_ok := FALSE;
	    END_IF;
	
	    IF ((#ars_statusword & 16#0800) = 16#0800)    //Bit 11 vom ZSW1
	        THEN #home_valid:= TRUE;
	        ELSE #home_valid:= FALSE;
	    END_IF;    
	
	    IF ((#ars_statusword & 16#0400) = 16#0400)    //Bit 10 vom ZSW1
	        THEN #pos_ok:= TRUE;
	        ELSE #pos_ok:= FALSE;
	    END_IF;    
	
	    IF ((#ars_statusword & 16#2000) = 16#2000)    //Bit 13 vom ZSW1
	        THEN #velo_zero:= TRUE;
	        ELSE #velo_zero:= FALSE;
	    END_IF;    
	
	    IF ((#ars_statusword & 16#0008) = 16#0008)    //Bit 3 vom ZSW1
	        THEN #fault:= TRUE;
	        ELSE #fault:= FALSE;
	    END_IF;    
	
	//************************************************************************************************
	
	//Schreiben Controlword
	
	 //  POKE (area := 16#84,
	 //        dbNumber := #DB_nr_position_word,
	 //        byteOffset := 2,
	 //        value := #ars_controlword );
	   
	    #A_Afag_soll_Werte.PROFIDRIVE_Controlword := #ars_controlword;
	    
	    
	    
	    
	    
END_FUNCTION_BLOCK

FUNCTION_BLOCK "BB_Ansteuerung_Afag_offen_V03.16"
TITLE = 'FB Positionierbetrieb'
{ S7_Optimized_Access := 'TRUE' }
AUTHOR : Essmann
FAMILY : metronix
NAME : position
VERSION : 1.1
//Der Baustein kann nicht rückübersetzt und unter STEP7 bearbeitet werden.  Der Baustein kann nur als Quelle im Ordner "Quellen" bearbeitet werden.    IO-Variablen  
   VAR_INPUT 
      E_UDT_Afag_ist_Werte : "Afag_ist_Werte";
      E_BA_Manuell : Bool;
      E_I_Manuell_Geschwindigkeit_Prozent : Int;
      E_Richten_reset_FRG : Bool;
      E_drive_enable : Bool := FALSE;
      E_start_homing : Bool := FALSE;
      E_abs_rel : Bool := FALSE;
      E_change_immediatly : Bool := FALSE;
      E_intermediate_stop : Bool := FALSE;
      E_hold : Bool := FALSE;
      E_jog_pos : Bool := FALSE;
      E_jog_neg : Bool := FALSE;
      E_fault_reset : Bool := FALSE;
      E_Tipp_pos : Bool;
      E_Tipp_neg : Bool;
      E_Start_pos_man : Bool;
      E_R_Verfahrweg_mm : Real;
      E_R_Afag_soll_wert_man_mm : Real;
      E_R_Softw_ES_min_mm : Real;
      E_R_Softw_ES_max_mm : Real;
      E_I_Max_Speed_mm_s : Int;
      E_I_Max_Beschleunigung_mm_s : Int;
   END_VAR

   VAR_OUTPUT 
      A_drive_enable_ok : Bool := FALSE;
      A_home_valid : Bool := FALSE;
      A_pos_ok : Bool := FALSE;
      A_velo_zero : Bool := FALSE;
      A_fault : Bool := FALSE;   // statische Variablen
      A_Positionsfehler : Bool;
      A_Fahrauftrag_Aktiv : Bool;
      A_Afag_ist_wert_mm : Real;
   END_VAR

   VAR_IN_OUT 
      E_A_UDT_Afag_Positionen : "Afag_Variablen_Positionen";
      A_UDT_Afag_soll_Werte : "Afag_soll_Werte";
   END_VAR

   VAR 
      switching_on_inhibited : Bool := FALSE;
      ready_for_switching_on : Bool := FALSE;
      switched_on : Bool := FALSE;
      operation : Bool := FALSE;
      ars_statusword : Word;
      ars_controlword : Word;
      start_pos : Bool := FALSE;
      start_pos_old : Bool := FALSE;   // ***********************************************************************************************************************Anweisungsteil
      start_pos_man : Bool;
      start_pos_man_old : Bool;
      Endlage_min_OK : Bool;
      Endlage_max_OK : Bool;
      Fahrauftrag_OK : Bool;
      AFAG_Ist_Wert_in_mm : Real;
      AFAG_soll_Wert_in_mm : Real;
      AFAG_soll_Speed_in_Prozent : Int;
      AFAG_soll_Beswchleunigung_in_mm_s : Int;
      R_TRIG_Instance {InstructionName := 'R_TRIG'; LibVersion := '1.0'} : R_TRIG;
      R_TRIG_Q_Tipp_neg : Bool;
      R_TRIG_Instance_1 {InstructionName := 'R_TRIG'; LibVersion := '1.0'} : R_TRIG;
      R_TRIG_Instance_2 {InstructionName := 'R_TRIG'; LibVersion := '1.0'} : R_TRIG;
      R_TRIG_Instance_3 {InstructionName := 'R_TRIG'; LibVersion := '1.0'} : R_TRIG;
      R_TRIG_Instance_4 {InstructionName := 'R_TRIG'; LibVersion := '1.0'} : R_TRIG;
      R_TRIG_Instance_5 {InstructionName := 'R_TRIG'; LibVersion := '1.0'} : R_TRIG;
      R_TRIG_Instance_6 {InstructionName := 'R_TRIG'; LibVersion := '1.0'} : R_TRIG;
      R_TRIG_Instance_7 {InstructionName := 'R_TRIG'; LibVersion := '1.0'} : R_TRIG;
      R_TRIG_Instance_8 {InstructionName := 'R_TRIG'; LibVersion := '1.0'} : R_TRIG;
      R_TRIG_Instance_9 {InstructionName := 'R_TRIG'; LibVersion := '1.0'} : R_TRIG;
      R_TRIG_Instance_10 {InstructionName := 'R_TRIG'; LibVersion := '1.0'} : R_TRIG;
      R_TRIG_Instance_11 {InstructionName := 'R_TRIG'; LibVersion := '1.0'} : R_TRIG;
      R_TRIG_Instance_12 {InstructionName := 'R_TRIG'; LibVersion := '1.0'} : R_TRIG;
      R_TRIG_Instance_13 {InstructionName := 'R_TRIG'; LibVersion := '1.0'} : R_TRIG;
      R_TRIG_Instance_14 {InstructionName := 'R_TRIG'; LibVersion := '1.0'} : R_TRIG;
      R_TRIG_Instance_15 {InstructionName := 'R_TRIG'; LibVersion := '1.0'} : R_TRIG;
      R_TRIG_Instance_16 {InstructionName := 'R_TRIG'; LibVersion := '1.0'} : R_TRIG;
      R_TRIG_Instance_17 {InstructionName := 'R_TRIG'; LibVersion := '1.0'} : R_TRIG;
      R_TRIG_Instance_18 {InstructionName := 'R_TRIG'; LibVersion := '1.0'} : R_TRIG;
   END_VAR


BEGIN
	
	
	//Ausgänge zuweisen
	#A_UDT_Afag_soll_Werte.Telegrammkennung := 16#e0;
	#A_Afag_ist_wert_mm := #AFAG_Ist_Wert_in_mm;
	#AFAG_Ist_Wert_in_mm := (DINT_TO_REAL(#E_UDT_Afag_ist_Werte.actual_position)) / 1.000000e+003;
	#A_UDT_Afag_soll_Werte.Zielposition := REAL_TO_DINT(#AFAG_soll_Wert_in_mm * 1.000000e+003);
	#A_UDT_Afag_soll_Werte.Fahrgeschwindigkeit := INT_TO_DINT(#AFAG_soll_Speed_in_Prozent * (#E_I_Max_Speed_mm_s / 100));
	#A_UDT_Afag_soll_Werte.Beschleunigung := INT_TO_DINT(#AFAG_soll_Beswchleunigung_in_mm_s);
	#E_A_UDT_Afag_Positionen.A_Softw_ES_min_mm := #E_R_Softw_ES_min_mm;
	#E_A_UDT_Afag_Positionen.A_Softw_ES_max_mm := #E_R_Softw_ES_max_mm;
	#E_A_UDT_Afag_Positionen.A_Max_Speed_mm_s := #E_I_Max_Speed_mm_s;
	#E_A_UDT_Afag_Positionen.A_Max_Beschleunigung_mm_s := #E_I_Max_Beschleunigung_mm_s;
	
	
	//************************************************************************************************
	
	//Lesen Statusword
	//Einlesen des Istzustands der Statemachine
	
	//    #DB_nr_actual_value_word:= INT_TO_WORD(#DB_nr_actual_value);
	//    #ars_statusword := PEEK_WORD (area := 16#84,
	//                                  dbNumber :=#DB_nr_actual_value_word,
	//                                  byteOffset := 2);
	#ars_statusword := #E_UDT_Afag_ist_Werte.PROFIDRIVE_Statusword;
	
	//Lesen Controlword
	//
	//  #DB_nr_position_word:=  INT_TO_WORD(#DB_nr_position);
	//  #ars_controlword := PEEK_WORD (area := 16#84,
	//                                  dbNumber :=#DB_nr_position_word,
	//                                  byteOffset := 2);
	
	// #ars_controlword := #A_UDT_Afag_soll_Werte.PROFIDRIVE_Controlword;
	
	//Steuern der Statemachine, S1 -> S2 -> S3 -> S4
	
	IF (#switching_on_inhibited                          //wenn state "switching_on_inhibited"
	    AND #E_drive_enable)                             //und  Reglerfreigabe
	THEN
	    #ars_controlword := 16#0406;              //dann state "ready_for_switching_on" anfordern,
	ELSIF (#switching_on_inhibited                     //
	    AND (NOT (#E_drive_enable)))                      //wenn Reglerfreigabe aus,
	THEN
	    #ars_controlword := 16#0400;              //dann state "switching_on_inhibited" anfordern.
	END_IF;
	
	IF (#ready_for_switching_on                          //wenn state "ready_for_switching_on"
	    AND #E_drive_enable)                             //und Reglerfeigabe
	THEN
	    #ars_controlword := 16#0407;              //dann state "switched_on" anfordern,
	ELSIF (#ready_for_switching_on                     //
	    AND (NOT (#E_drive_enable)))                      //wenn Reglerfeigabe aus,
	THEN
	    #ars_controlword := 16#0400;              //dann state "switching_on_inhibited" anfordern.
	END_IF;
	
	IF (#switched_on                                     //wenn state "switched_on"
	    AND #E_drive_enable)                             //und Reglerfeigabe
	THEN
	    #ars_controlword := 16#040f;              //dann state "operation" anfordern,
	ELSIF (#switched_on                                //
	    AND (NOT (#E_drive_enable)))                      //wenn Reglerfeigabe aus,
	THEN
	    #ars_controlword := 16#0400;              //dann state "switching_on_inhibited" anfordern.
	END_IF;
	
	IF (#operation                                       //wenn state "operation"
	    AND (NOT (#E_drive_enable)))                      //und keine Reglerfeigabe
	THEN
	    #ars_controlword := 16#040e;              //dann state "switching_on_inhibited" anfordern.
	END_IF;
	
	//************************************************************************************************
	
	//Kommandos über digitale Eingänge
	// Bit 10 (control by plc) im Controlword muss immer gesetzt sein
	
	IF #E_start_homing
	THEN
	    #ars_controlword := (#ars_controlword OR 16#0C00);    //Setzen Bit 11 im STW1
	ELSE
	    #ars_controlword := (#ars_controlword & 16#f7ff);
	END_IF;
	
	IF (#Fahrauftrag_OK = 1) THEN
	    IF (#start_pos_old <> #start_pos) OR (#start_pos_man_old <> #start_pos_man)
	    THEN
	        IF #start_pos OR #start_pos_man
	        THEN
	            #ars_controlword := (#ars_controlword OR 16#0440);    //Setzen Bit 6 im STW1
	        ELSE
	            #ars_controlword := (#ars_controlword & 16#ffbf);
	        END_IF;
	    END_IF;
	    
	    #start_pos_old := #start_pos;
	    #start_pos_man_old := #start_pos_man;
	    
	END_IF;
	
	
	IF #E_abs_rel
	THEN
	    #ars_controlword := (#ars_controlword OR 16#1400);   //Setzen Bit 12 im STW1
	ELSE
	    #ars_controlword := (#ars_controlword & 16#efff);
	END_IF;
	
	IF #E_change_immediatly
	THEN
	    #ars_controlword := (#ars_controlword OR 16#2400);   //Setzen Bit 13 im STW1
	ELSE
	    #ars_controlword := (#ars_controlword & 16#dfff);
	END_IF;
	
	IF #E_intermediate_stop
	THEN
	    #ars_controlword := (#ars_controlword & 16#ffdf);   //Rücksetzen Bit 5 im STW1
	ELSE
	    #ars_controlword := (#ars_controlword OR 16#0420);
	END_IF;
	
	IF #E_hold
	THEN
	    #ars_controlword := (#ars_controlword & 16#ffef);    //Rücksetzen Bit 4 im STW1
	    #ars_controlword := (#ars_controlword & 16#feff);    //Rücksetzen jog_pos
	    #ars_controlword := (#ars_controlword & 16#fdff);    //Rücksetzen jog_neg
	ELSE
	    #ars_controlword := (#ars_controlword OR 16#0410);
	END_IF;
	
	IF (#E_jog_pos AND NOT #E_hold) AND (#AFAG_Ist_Wert_in_mm < #E_R_Softw_ES_max_mm)
	THEN
	    #ars_controlword := (#ars_controlword OR 16#0500);    //Setzen Bit 8 im STW1
	ELSE
	    #ars_controlword := (#ars_controlword & 16#feff);
	END_IF;
	
	IF (#E_jog_neg AND NOT #E_hold) AND (#AFAG_Ist_Wert_in_mm > #E_R_Softw_ES_min_mm)
	THEN
	    #ars_controlword := (#ars_controlword OR 16#0600);    //Setzen Bit 9 im STW1
	ELSE
	    #ars_controlword := (#ars_controlword & 16#fdff);
	END_IF;
	
	IF #E_fault_reset
	THEN
	    #ars_controlword := (#ars_controlword OR 16#0480);    //Setzen Bit 7 im STW1
	ELSE
	    #ars_controlword := (#ars_controlword & 16#ff7f);
	END_IF;
	
	
	//************************************************************************************************
	
	//Setzen digitaler Ausgänge
	
	IF #operation
	THEN
	    #A_drive_enable_ok := TRUE;
	ELSE
	    #A_drive_enable_ok := FALSE;
	END_IF;
	
	IF ((#ars_statusword & 16#0800) = 16#0800)    //Bit 11 vom ZSW1
	THEN
	    #A_home_valid := TRUE;
	ELSE
	    #A_home_valid := FALSE;
	END_IF;
	
	IF ((#ars_statusword & 16#0400) = 16#0400)    //Bit 10 vom ZSW1
	THEN
	    #A_pos_ok := TRUE;
	ELSE
	    #A_pos_ok := FALSE;
	END_IF;
	
	IF ((#ars_statusword & 16#2000) = 16#2000)    //Bit 13 vom ZSW1
	THEN
	    #A_velo_zero := TRUE;
	ELSE
	    #A_velo_zero := FALSE;
	END_IF;
	
	IF ((#ars_statusword & 16#0008) = 16#0008)    //Bit 3 vom ZSW1
	THEN
	    #A_fault := TRUE;
	ELSE
	    #A_fault := FALSE;
	END_IF;
	
	//************************************************************************************************
	
	//Schreiben Controlword
	
	//  POKE (area := 16#84,
	//        dbNumber := #DB_nr_position_word,
	//        byteOffset := 2,
	//        value := #ars_controlword );
	
	#A_UDT_Afag_soll_Werte.PROFIDRIVE_Controlword := #ars_controlword;
	
	
	
	
	
	
	// Achse mit Position Starten
	// Position[0]
	#R_TRIG_Instance_3(CLK := #E_A_UDT_Afag_Positionen.Start_POS_Position[0]);
	IF #R_TRIG_Instance_3.Q THEN
	    #AFAG_soll_Wert_in_mm := #E_A_UDT_Afag_Positionen.Soll_Wert_in_mm_Position[0];
	    #AFAG_soll_Beswchleunigung_in_mm_s := #E_A_UDT_Afag_Positionen.Soll_Beschleunigung_in_mm_s_Position[0];
	    #start_pos := true;
	    
	    #AFAG_soll_Speed_in_Prozent := #E_A_UDT_Afag_Positionen.Soll_Speed_in_Prozent_Position[0];
	END_IF;
	
	// Position[1]
	#R_TRIG_Instance_4(CLK:=#E_A_UDT_Afag_Positionen.Start_POS_Position[1]);
	IF #R_TRIG_Instance_4.Q THEN
	    #AFAG_soll_Wert_in_mm := #E_A_UDT_Afag_Positionen.Soll_Wert_in_mm_Position[1];
	    #AFAG_soll_Beswchleunigung_in_mm_s := #E_A_UDT_Afag_Positionen.Soll_Beschleunigung_in_mm_s_Position[1];
	    #start_pos := true;
	
	    #AFAG_soll_Speed_in_Prozent := #E_A_UDT_Afag_Positionen.Soll_Speed_in_Prozent_Position[1];
	END_IF;
	
	
	// Position 2
	#R_TRIG_Instance_5(CLK:=#E_A_UDT_Afag_Positionen.Start_POS_Position[2]);
	IF #R_TRIG_Instance_5.Q THEN
	    #AFAG_soll_Wert_in_mm := #E_A_UDT_Afag_Positionen.Soll_Wert_in_mm_Position[2];
	    #AFAG_soll_Beswchleunigung_in_mm_s := #E_A_UDT_Afag_Positionen.Soll_Beschleunigung_in_mm_s_Position[2];
	    #start_pos := true;
	
	    #AFAG_soll_Speed_in_Prozent := #E_A_UDT_Afag_Positionen.Soll_Speed_in_Prozent_Position[2];
	END_IF;
	
	// Position 3
	#R_TRIG_Instance_6(CLK := #E_A_UDT_Afag_Positionen.Start_POS_Position[3]);
	IF #R_TRIG_Instance_6.Q THEN
	    #AFAG_soll_Wert_in_mm := #E_A_UDT_Afag_Positionen.Soll_Wert_in_mm_Position[3];
	    #AFAG_soll_Beswchleunigung_in_mm_s := #E_A_UDT_Afag_Positionen.Soll_Beschleunigung_in_mm_s_Position[3];
	    #start_pos := true;
	
	    #AFAG_soll_Speed_in_Prozent := #E_A_UDT_Afag_Positionen.Soll_Speed_in_Prozent_Position[3];
	END_IF;
	
	// Position 4
	#R_TRIG_Instance_7(CLK := #E_A_UDT_Afag_Positionen.Start_POS_Position[4]);
	IF #R_TRIG_Instance_7.Q THEN
	    #AFAG_soll_Wert_in_mm := #E_A_UDT_Afag_Positionen.Soll_Wert_in_mm_Position[4];
	    #AFAG_soll_Beswchleunigung_in_mm_s := #E_A_UDT_Afag_Positionen.Soll_Beschleunigung_in_mm_s_Position[4];
	    #start_pos := true;
	
	    #AFAG_soll_Speed_in_Prozent := #E_A_UDT_Afag_Positionen.Soll_Speed_in_Prozent_Position[4];
	END_IF;
	
	// Position 5
	#R_TRIG_Instance_8(CLK := #E_A_UDT_Afag_Positionen.Start_POS_Position[5]);
	IF #R_TRIG_Instance_8.Q THEN
	    #AFAG_soll_Wert_in_mm := #E_A_UDT_Afag_Positionen.Soll_Wert_in_mm_Position[5];
	    #AFAG_soll_Beswchleunigung_in_mm_s := #E_A_UDT_Afag_Positionen.Soll_Beschleunigung_in_mm_s_Position[5];
	    #start_pos := true;
	
	    #AFAG_soll_Speed_in_Prozent := #E_A_UDT_Afag_Positionen.Soll_Speed_in_Prozent_Position[5];
	END_IF;
	
	// Position 6
	#R_TRIG_Instance_9(CLK := #E_A_UDT_Afag_Positionen.Start_POS_Position[6]);
	IF #R_TRIG_Instance_9.Q THEN
	    #AFAG_soll_Wert_in_mm := #E_A_UDT_Afag_Positionen.Soll_Wert_in_mm_Position[6];
	    #AFAG_soll_Beswchleunigung_in_mm_s := #E_A_UDT_Afag_Positionen.Soll_Beschleunigung_in_mm_s_Position[6];
	    #start_pos := true;
	
	    #AFAG_soll_Speed_in_Prozent := #E_A_UDT_Afag_Positionen.Soll_Speed_in_Prozent_Position[6];
	END_IF;
	
	// Position 7
	#R_TRIG_Instance_10(CLK := #E_A_UDT_Afag_Positionen.Start_POS_Position[7]);
	IF #R_TRIG_Instance_10.Q THEN
	    #AFAG_soll_Wert_in_mm := #E_A_UDT_Afag_Positionen.Soll_Wert_in_mm_Position[7];
	    #AFAG_soll_Beswchleunigung_in_mm_s := #E_A_UDT_Afag_Positionen.Soll_Beschleunigung_in_mm_s_Position[7];
	    #start_pos := true;
	
	    #AFAG_soll_Speed_in_Prozent := #E_A_UDT_Afag_Positionen.Soll_Speed_in_Prozent_Position[7];
	END_IF;
	
	// Position 8
	#R_TRIG_Instance_11(CLK := #E_A_UDT_Afag_Positionen.Start_POS_Position[8]);
	IF #R_TRIG_Instance_11.Q THEN
	    #AFAG_soll_Wert_in_mm := #E_A_UDT_Afag_Positionen.Soll_Wert_in_mm_Position[8];
	    #AFAG_soll_Beswchleunigung_in_mm_s := #E_A_UDT_Afag_Positionen.Soll_Beschleunigung_in_mm_s_Position[8];
	    #start_pos := true;
	
	    #AFAG_soll_Speed_in_Prozent := #E_A_UDT_Afag_Positionen.Soll_Speed_in_Prozent_Position[8];
	END_IF;
	
	// Position 9
	#R_TRIG_Instance_12(CLK := #E_A_UDT_Afag_Positionen.Start_POS_Position[9]);
	IF #R_TRIG_Instance_12.Q THEN
	    #AFAG_soll_Wert_in_mm := #E_A_UDT_Afag_Positionen.Soll_Wert_in_mm_Position[9];
	    #AFAG_soll_Beswchleunigung_in_mm_s := #E_A_UDT_Afag_Positionen.Soll_Beschleunigung_in_mm_s_Position[9];
	    #start_pos := true;
	
	    #AFAG_soll_Speed_in_Prozent := #E_A_UDT_Afag_Positionen.Soll_Speed_in_Prozent_Position[9];
	END_IF;
	
	// Position 10
	#R_TRIG_Instance_13(CLK := #E_A_UDT_Afag_Positionen.Start_POS_Position[10]);
	IF #R_TRIG_Instance_13.Q THEN
	    #AFAG_soll_Wert_in_mm := #E_A_UDT_Afag_Positionen.Soll_Wert_in_mm_Position[10];
	    #AFAG_soll_Beswchleunigung_in_mm_s := #E_A_UDT_Afag_Positionen.Soll_Beschleunigung_in_mm_s_Position[10];
	    #start_pos := true;
	
	    #AFAG_soll_Speed_in_Prozent := #E_A_UDT_Afag_Positionen.Soll_Speed_in_Prozent_Position[10];
	END_IF;
	
	// Position 11
	#R_TRIG_Instance_14(CLK := #E_A_UDT_Afag_Positionen.Start_POS_Position[11]);
	IF #R_TRIG_Instance_14.Q THEN
	    #AFAG_soll_Wert_in_mm := #E_A_UDT_Afag_Positionen.Soll_Wert_in_mm_Position[11];
	    #AFAG_soll_Beswchleunigung_in_mm_s := #E_A_UDT_Afag_Positionen.Soll_Beschleunigung_in_mm_s_Position[11];
	    #start_pos := true;
	
	    #AFAG_soll_Speed_in_Prozent := #E_A_UDT_Afag_Positionen.Soll_Speed_in_Prozent_Position[11];
	END_IF;
	
	// Position 12
	#R_TRIG_Instance_15(CLK := #E_A_UDT_Afag_Positionen.Start_POS_Position[12]);
	IF #R_TRIG_Instance_15.Q THEN
	    #AFAG_soll_Wert_in_mm := #E_A_UDT_Afag_Positionen.Soll_Wert_in_mm_Position[12];
	    #AFAG_soll_Beswchleunigung_in_mm_s := #E_A_UDT_Afag_Positionen.Soll_Beschleunigung_in_mm_s_Position[12];
	    #start_pos := true;
	
	    #AFAG_soll_Speed_in_Prozent := #E_A_UDT_Afag_Positionen.Soll_Speed_in_Prozent_Position[12];
	END_IF;
	
	// Position 13
	#R_TRIG_Instance_16(CLK := #E_A_UDT_Afag_Positionen.Start_POS_Position[13]);
	IF #R_TRIG_Instance_16.Q THEN
	    #AFAG_soll_Wert_in_mm := #E_A_UDT_Afag_Positionen.Soll_Wert_in_mm_Position[13];
	    #AFAG_soll_Beswchleunigung_in_mm_s := #E_A_UDT_Afag_Positionen.Soll_Beschleunigung_in_mm_s_Position[13];
	    #start_pos := true;
	
	    #AFAG_soll_Speed_in_Prozent := #E_A_UDT_Afag_Positionen.Soll_Speed_in_Prozent_Position[13];
	END_IF;
	
	// Position 14
	#R_TRIG_Instance_17(CLK := #E_A_UDT_Afag_Positionen.Start_POS_Position[14]);
	IF #R_TRIG_Instance_17.Q THEN
	    #AFAG_soll_Wert_in_mm := #E_A_UDT_Afag_Positionen.Soll_Wert_in_mm_Position[14];
	    #AFAG_soll_Beswchleunigung_in_mm_s := #E_A_UDT_Afag_Positionen.Soll_Beschleunigung_in_mm_s_Position[14];
	    #start_pos := true;
	
	    #AFAG_soll_Speed_in_Prozent := #E_A_UDT_Afag_Positionen.Soll_Speed_in_Prozent_Position[14];
	END_IF;
	
	// Position 15
	#R_TRIG_Instance_18(CLK:= #E_A_UDT_Afag_Positionen.Start_POS_Position[15]);
	IF #R_TRIG_Instance_18.Q THEN
	    #AFAG_soll_Wert_in_mm := #E_A_UDT_Afag_Positionen.Soll_Wert_in_mm_Position[15];
	    #AFAG_soll_Beswchleunigung_in_mm_s := #E_A_UDT_Afag_Positionen.Soll_Beschleunigung_in_mm_s_Position[15];
	    #start_pos := true;
	   
	    #AFAG_soll_Speed_in_Prozent := #E_A_UDT_Afag_Positionen.Soll_Speed_in_Prozent_Position[15];
	END_IF;
	
	//Manuelle Geschwindigkeitsanpassung
	IF #E_BA_Manuell = TRUE THEN
	    #AFAG_soll_Speed_in_Prozent := #E_I_Manuell_Geschwindigkeit_Prozent;
	    #AFAG_soll_Beswchleunigung_in_mm_s := 100;
	END_IF;
	
	IF( (#E_A_UDT_Afag_Positionen.Start_POS_Position[0] AND #E_A_UDT_Afag_Positionen.POS_OK_Position[0])OR
	   (#E_A_UDT_Afag_Positionen.Start_POS_Position[1]AND #E_A_UDT_Afag_Positionen.POS_OK_Position[1])OR
	   (#E_A_UDT_Afag_Positionen.Start_POS_Position[2]AND #E_A_UDT_Afag_Positionen.POS_OK_Position[2])OR
	   (#E_A_UDT_Afag_Positionen.Start_POS_Position[3]AND #E_A_UDT_Afag_Positionen.POS_OK_Position[3])OR
	   (#E_A_UDT_Afag_Positionen.Start_POS_Position[4]AND #E_A_UDT_Afag_Positionen.POS_OK_Position[4])OR
	   (#E_A_UDT_Afag_Positionen.Start_POS_Position[5]AND #E_A_UDT_Afag_Positionen.POS_OK_Position[5])OR
	   (#E_A_UDT_Afag_Positionen.Start_POS_Position[6]AND #E_A_UDT_Afag_Positionen.POS_OK_Position[6])OR
	   (#E_A_UDT_Afag_Positionen.Start_POS_Position[7]AND #E_A_UDT_Afag_Positionen.POS_OK_Position[7])OR
	   (#E_A_UDT_Afag_Positionen.Start_POS_Position[8]AND #E_A_UDT_Afag_Positionen.POS_OK_Position[8])OR
	   (#E_A_UDT_Afag_Positionen.Start_POS_Position[9]AND #E_A_UDT_Afag_Positionen.POS_OK_Position[9])OR
	   (#E_A_UDT_Afag_Positionen.Start_POS_Position[10]AND #E_A_UDT_Afag_Positionen.POS_OK_Position[10])OR
	   (#E_A_UDT_Afag_Positionen.Start_POS_Position[11]AND #E_A_UDT_Afag_Positionen.POS_OK_Position[11])OR
	   (#E_A_UDT_Afag_Positionen.Start_POS_Position[12]AND #E_A_UDT_Afag_Positionen.POS_OK_Position[12])OR
	   (#E_A_UDT_Afag_Positionen.Start_POS_Position[13]AND #E_A_UDT_Afag_Positionen.POS_OK_Position[13])OR
	   (#E_A_UDT_Afag_Positionen.Start_POS_Position[14]AND #E_A_UDT_Afag_Positionen.POS_OK_Position[14])OR
	   (#E_A_UDT_Afag_Positionen.Start_POS_Position[15]AND #E_A_UDT_Afag_Positionen.POS_OK_Position[15])OR
	    #A_Positionsfehler OR #E_Richten_reset_FRG)
	THEN
	    #start_pos := 0;
	    #E_A_UDT_Afag_Positionen.Start_POS_Position[0] := 0;
	    #E_A_UDT_Afag_Positionen.Start_POS_Position[1] := 0;
	    #E_A_UDT_Afag_Positionen.Start_POS_Position[2] := 0;
	    #E_A_UDT_Afag_Positionen.Start_POS_Position[3] := 0;
	    #E_A_UDT_Afag_Positionen.Start_POS_Position[4] := 0;
	    #E_A_UDT_Afag_Positionen.Start_POS_Position[5] := 0;
	    #E_A_UDT_Afag_Positionen.Start_POS_Position[6] := 0;
	    #E_A_UDT_Afag_Positionen.Start_POS_Position[7] := 0;
	    #E_A_UDT_Afag_Positionen.Start_POS_Position[8] := 0;
	    #E_A_UDT_Afag_Positionen.Start_POS_Position[9] := 0;
	    #E_A_UDT_Afag_Positionen.Start_POS_Position[10] := 0;
	    #E_A_UDT_Afag_Positionen.Start_POS_Position[11] := 0;
	    #E_A_UDT_Afag_Positionen.Start_POS_Position[12] := 0;
	    #E_A_UDT_Afag_Positionen.Start_POS_Position[13] := 0;
	    #E_A_UDT_Afag_Positionen.Start_POS_Position[14] := 0;
	    #E_A_UDT_Afag_Positionen.Start_POS_Position[15] := 0;
	    #E_A_UDT_Afag_Positionen.POS_OK_Position[15] := 0;
	END_IF;
	
	
	// Achse Positionsrückmeldung
	
	IF ((ABS(#AFAG_Ist_Wert_in_mm - #E_A_UDT_Afag_Positionen.Soll_Wert_in_mm_Position[0])) < #E_A_UDT_Afag_Positionen.Positionstoleranz_Position[0])
	THEN
	    #E_A_UDT_Afag_Positionen.POS_OK_Position[0] := 1;
	ELSE
	    #E_A_UDT_Afag_Positionen.POS_OK_Position[0] := 0;
	END_IF;
	
	IF ((ABS(#AFAG_Ist_Wert_in_mm - #E_A_UDT_Afag_Positionen.Soll_Wert_in_mm_Position[1])) < #E_A_UDT_Afag_Positionen.Positionstoleranz_Position[1])
	THEN
	    #E_A_UDT_Afag_Positionen.POS_OK_Position[1] := 1;
	ELSE
	    #E_A_UDT_Afag_Positionen.POS_OK_Position[1] := 0;
	END_IF;
	
	IF ((ABS(#AFAG_Ist_Wert_in_mm - #E_A_UDT_Afag_Positionen.Soll_Wert_in_mm_Position[2])) < #E_A_UDT_Afag_Positionen.Positionstoleranz_Position[2])
	THEN
	    #E_A_UDT_Afag_Positionen.POS_OK_Position[2] := 1;
	ELSE
	    #E_A_UDT_Afag_Positionen.POS_OK_Position[2] := 0;
	END_IF;
	
	IF ((ABS(#AFAG_Ist_Wert_in_mm - #E_A_UDT_Afag_Positionen.Soll_Wert_in_mm_Position[3])) < #E_A_UDT_Afag_Positionen.Positionstoleranz_Position[3])
	THEN
	    #E_A_UDT_Afag_Positionen.POS_OK_Position[3] := 1;
	ELSE
	    #E_A_UDT_Afag_Positionen.POS_OK_Position[3] := 0;
	END_IF;
	
	IF ((ABS(#AFAG_Ist_Wert_in_mm - #E_A_UDT_Afag_Positionen.Soll_Wert_in_mm_Position[4])) < #E_A_UDT_Afag_Positionen.Positionstoleranz_Position[4])
	THEN
	    #E_A_UDT_Afag_Positionen.POS_OK_Position[4] := 1;
	ELSE
	    #E_A_UDT_Afag_Positionen.POS_OK_Position[4] := 0;
	END_IF;
	
	IF ((ABS(#AFAG_Ist_Wert_in_mm - #E_A_UDT_Afag_Positionen.Soll_Wert_in_mm_Position[5])) < #E_A_UDT_Afag_Positionen.Positionstoleranz_Position[5])
	THEN
	    #E_A_UDT_Afag_Positionen.POS_OK_Position[5] := 1;
	ELSE
	    #E_A_UDT_Afag_Positionen.POS_OK_Position[5] := 0;
	END_IF;
	
	IF ((ABS(#AFAG_Ist_Wert_in_mm - #E_A_UDT_Afag_Positionen.Soll_Wert_in_mm_Position[6])) < #E_A_UDT_Afag_Positionen.Positionstoleranz_Position[6])
	THEN
	    #E_A_UDT_Afag_Positionen.POS_OK_Position[6] := 1;
	ELSE
	    #E_A_UDT_Afag_Positionen.POS_OK_Position[6] := 0;
	END_IF;
	
	IF ((ABS(#AFAG_Ist_Wert_in_mm - #E_A_UDT_Afag_Positionen.Soll_Wert_in_mm_Position[7])) < #E_A_UDT_Afag_Positionen.Positionstoleranz_Position[7])
	THEN
	    #E_A_UDT_Afag_Positionen.POS_OK_Position[7] := 1;
	ELSE
	    #E_A_UDT_Afag_Positionen.POS_OK_Position[7] := 0;
	END_IF;
	
	IF ((ABS(#AFAG_Ist_Wert_in_mm - #E_A_UDT_Afag_Positionen.Soll_Wert_in_mm_Position[8])) < #E_A_UDT_Afag_Positionen.Positionstoleranz_Position[8])
	THEN
	    #E_A_UDT_Afag_Positionen.POS_OK_Position[8] := 1;
	ELSE
	    #E_A_UDT_Afag_Positionen.POS_OK_Position[8] := 0;
	END_IF;
	
	IF ((ABS(#AFAG_Ist_Wert_in_mm - #E_A_UDT_Afag_Positionen.Soll_Wert_in_mm_Position[9])) < #E_A_UDT_Afag_Positionen.Positionstoleranz_Position[9])
	THEN
	    #E_A_UDT_Afag_Positionen.POS_OK_Position[9] := 1;
	ELSE
	    #E_A_UDT_Afag_Positionen.POS_OK_Position[9] := 0;
	END_IF;
	
	IF ((ABS(#AFAG_Ist_Wert_in_mm - #E_A_UDT_Afag_Positionen.Soll_Wert_in_mm_Position[10])) < #E_A_UDT_Afag_Positionen.Positionstoleranz_Position[10])
	THEN
	    #E_A_UDT_Afag_Positionen.POS_OK_Position[10] := 1;
	ELSE
	    #E_A_UDT_Afag_Positionen.POS_OK_Position[10] := 0;
	END_IF;
	
	IF ((ABS(#AFAG_Ist_Wert_in_mm - #E_A_UDT_Afag_Positionen.Soll_Wert_in_mm_Position[11])) < #E_A_UDT_Afag_Positionen.Positionstoleranz_Position[11])
	THEN
	    #E_A_UDT_Afag_Positionen.POS_OK_Position[11] := 1;
	ELSE
	    #E_A_UDT_Afag_Positionen.POS_OK_Position[11] := 0;
	END_IF;
	
	IF ((ABS(#AFAG_Ist_Wert_in_mm - #E_A_UDT_Afag_Positionen.Soll_Wert_in_mm_Position[12])) < #E_A_UDT_Afag_Positionen.Positionstoleranz_Position[12])
	THEN
	    #E_A_UDT_Afag_Positionen.POS_OK_Position[12] := 1;
	ELSE
	    #E_A_UDT_Afag_Positionen.POS_OK_Position[12] := 0;
	END_IF;
	
	IF ((ABS(#AFAG_Ist_Wert_in_mm - #E_A_UDT_Afag_Positionen.Soll_Wert_in_mm_Position[13])) < #E_A_UDT_Afag_Positionen.Positionstoleranz_Position[13])
	THEN
	    #E_A_UDT_Afag_Positionen.POS_OK_Position[13] := 1;
	ELSE
	    #E_A_UDT_Afag_Positionen.POS_OK_Position[13] := 0;
	END_IF;
	
	IF ((ABS(#AFAG_Ist_Wert_in_mm - #E_A_UDT_Afag_Positionen.Soll_Wert_in_mm_Position[14])) < #E_A_UDT_Afag_Positionen.Positionstoleranz_Position[14])
	THEN
	    #E_A_UDT_Afag_Positionen.POS_OK_Position[14] := 1;
	ELSE
	    #E_A_UDT_Afag_Positionen.POS_OK_Position[14] := 0;
	END_IF;
	
	IF ((ABS(#AFAG_Ist_Wert_in_mm - #E_A_UDT_Afag_Positionen.Soll_Wert_in_mm_Position[15])) < #E_A_UDT_Afag_Positionen.Positionstoleranz_Position[15])
	THEN
	    #E_A_UDT_Afag_Positionen.POS_OK_Position[15] := 1;
	ELSE
	    #E_A_UDT_Afag_Positionen.POS_OK_Position[15] := 0;
	END_IF;
	
	IF
	    (#E_A_UDT_Afag_Positionen.Start_POS_Position[0]) OR
	    (#E_A_UDT_Afag_Positionen.Start_POS_Position[1]) OR
	    (#E_A_UDT_Afag_Positionen.Start_POS_Position[2]) OR
	    (#E_A_UDT_Afag_Positionen.Start_POS_Position[3]) OR
	    (#E_A_UDT_Afag_Positionen.Start_POS_Position[4]) OR
	    (#E_A_UDT_Afag_Positionen.Start_POS_Position[5]) OR
	    (#E_A_UDT_Afag_Positionen.Start_POS_Position[6]) OR
	    (#E_A_UDT_Afag_Positionen.Start_POS_Position[7]) OR
	    (#E_A_UDT_Afag_Positionen.Start_POS_Position[8]) OR
	    (#E_A_UDT_Afag_Positionen.Start_POS_Position[9]) OR
	    (#E_A_UDT_Afag_Positionen.Start_POS_Position[10]) OR
	    (#E_A_UDT_Afag_Positionen.Start_POS_Position[11]) OR
	    (#E_A_UDT_Afag_Positionen.Start_POS_Position[12]) OR
	    (#E_A_UDT_Afag_Positionen.Start_POS_Position[13]) OR
	    (#E_A_UDT_Afag_Positionen.Start_POS_Position[14]) OR
	    (#E_A_UDT_Afag_Positionen.Start_POS_Position[15]) OR
	    (#start_pos)
	THEN
	    #A_Fahrauftrag_Aktiv := 1;
	ELSE
	    #A_Fahrauftrag_Aktiv := 0;
	END_IF;
	
	
	
	
	//Reset Start pos
	IF ((#A_pos_ok = true) OR (#A_drive_enable_ok = FALSE) OR (#E_fault_reset = TRUE))
	THEN
	    #start_pos_man := false;
	END_IF;
	
	//Tipp pos
	#R_TRIG_Instance(CLK:=#E_Tipp_pos);
	IF (#R_TRIG_Instance.Q AND NOT #start_pos_man)
	THEN
	    #AFAG_soll_Wert_in_mm := #AFAG_Ist_Wert_in_mm + #E_R_Verfahrweg_mm;
	    #start_pos_man := TRUE;
	END_IF;
	
	//Tipp neg
	#R_TRIG_Instance_1(CLK:=#E_Tipp_neg);
	IF (#R_TRIG_Instance_1.Q AND NOT #start_pos_man)
	THEN
	    #AFAG_soll_Wert_in_mm := #AFAG_Ist_Wert_in_mm - #E_R_Verfahrweg_mm;
	    #start_pos_man := TRUE;
	END_IF;
	
	//absolut verfahren
	#R_TRIG_Instance_2(CLK:=#E_Start_pos_man);
	IF(#R_TRIG_Instance_2.Q AND NOT #start_pos_man)
	THEN
	    #AFAG_soll_Wert_in_mm := #E_R_Afag_soll_wert_man_mm;
	    #start_pos_man := TRUE;
	END_IF;
	
	// Endlagen Überwachen
	IF (#AFAG_Ist_Wert_in_mm > #E_R_Softw_ES_min_mm)
	THEN
	    #Endlage_min_OK := TRUE;
	ELSE
	    #Endlage_min_OK := FALSE;
	END_IF;
	
	IF (#AFAG_Ist_Wert_in_mm < #E_R_Softw_ES_max_mm)
	THEN
	    #Endlage_max_OK := TRUE;
	ELSE
	    #Endlage_max_OK := FALSE;
	END_IF;
	
	//Überwachung Fahrauftrag
	IF (#Endlage_min_OK AND #Endlage_max_OK)
	THEN
	    #Fahrauftrag_OK := TRUE;
	ELSE
	    #Fahrauftrag_OK := FALSE;
	END_IF;
	
	//Störmeldung Positionierung
	IF (#Endlage_min_OK AND #Endlage_max_OK AND #Fahrauftrag_OK)
	THEN
	    #A_Positionsfehler := FALSE;
	ELSE
	    #A_Positionsfehler := TRUE;
	END_IF;
	    
	//Einlesen des Istzustands der Statemachine
	   IF ((#ars_statusword & 16#0047) = 16#0040)
	        THEN #switching_on_inhibited := TRUE;
	        ELSE #switching_on_inhibited := FALSE;
	    END_IF;
	
	    IF ((#ars_statusword & 16#0047) = 16#0001)
	        THEN #ready_for_switching_on:= TRUE;
	        ELSE #ready_for_switching_on:= FALSE;
	    END_IF;
	     
	    IF ((#ars_statusword & 16#0047) = 16#0003)
	        THEN #switched_on:= TRUE;
	        ELSE #switched_on:= FALSE;
	    END_IF;
	
	    IF ((#ars_statusword & 16#0047) = 16#0007)
	        THEN #operation:= TRUE;
	        ELSE #operation:= FALSE;
	    END_IF;    
	
	
	
	    
	    
END_FUNCTION_BLOCK

FUNCTION_BLOCK "Drehtelleransteuerung_SCL"
{ S7_Optimized_Access := 'TRUE' }
VERSION : 0.1
   VAR_INPUT RETAIN
      ES_in_Position : Bool;
      ES_Motor_aus : Bool;
      Motorschutz : Bool;
      Automatik : Bool;
      Manuell : Bool;
      Ablauf_aktiv : Bool;
      Richten : Bool;
      SM_reset : Bool;
      Reset_Frg : Bool;
      Not_Aus_OK : Bool;
      Tueren_OK : Bool;
      Lichtvorhang_OK : Bool;
      Sicherheitsbit_DT : Bool;
      TP_Taste_tippen : Bool;
      Start_taste_tippen : Bool;
      links0_rechts1_drehen : Bool;
      Time_Drehteller_Laufzeit : Time;
      Time_Drehteller_nicht_in_Position : Time;
      Time_Öffnungszeit_Bremse : Time;
      Time_Startzeit : Time;
      Wartungsintervall : DInt;
   END_VAR

   VAR_OUTPUT RETAIN
      Schuetz_links : Bool;
      Schuetz_rechts : Bool;
      DT_Bremse : Bool;
      Aktorzyklen : DInt;
   END_VAR

   VAR_IN_OUT RETAIN
      Freigabe_DT : Bool;
      Manuellfreigabe : Bool;
      Richtenfreigabe : Bool;
      Fertigmeldung_Drehteller : Bool;
      Betriebsfertigmeldung : Bool;
      SM_Drehteller_dreht_nicht : Bool;
      SM_Drehteller_nicht_in_Position : Bool;
      SM_Motorschutz : Bool;
      SM_Sicherheitsbit : Bool;
      SM_Wartung : Bool;
   END_VAR
   VAR_IN_OUT DB_SPECIFIC
      Auto_Frg_Drehen_Vorwärts : Bool;
      Auto_Frg_Drehen_Rückwärts : Bool;
      Manu_Frg_Drehen_Vorwärts : Bool;
      Manu_Frg_Drehen_Rückwärts : Bool;
      Richt_Frg_Drehen_Vorwärts : Bool;
      Richt_Frg_Drehen_Rückwärts : Bool;
   END_VAR

   VAR RETAIN
      iStep : Int;
      Schrittkette_start : Bool;
      Befehlsfreigabe : Bool;
      Modolo_Wartungszähler : DInt;
      Timer_Drehteller_Laufzeit {InstructionName := 'TON_TIME'; LibVersion := '1.0'; S7_SetPoint := 'False'} : TON_TIME;
      Timer_Drehteller_nicht_in_Position {InstructionName := 'TON_TIME'; LibVersion := '1.0'; S7_SetPoint := 'False'} : TON_TIME;
   END_VAR
   VAR 
      F_TRIG_Zyklenzähler {InstructionName := 'F_TRIG'; LibVersion := '1.0'} : F_TRIG;
      F_TRIG_Modolo_gleich_0 {InstructionName := 'F_TRIG'; LibVersion := '1.0'} : F_TRIG;
   END_VAR
   VAR DB_SPECIFIC
      Timer_Öffnungszeit_Bremse {InstructionName := 'TON_TIME'; LibVersion := '1.0'; S7_SetPoint := 'False'} : TON_TIME;
      Timer_Startzeit {InstructionName := 'TON_TIME'; LibVersion := '1.0'; S7_SetPoint := 'False'} : TON_TIME;
      Temp_Vorwärts { ExternalAccessible := 'False'; ExternalVisible := 'False'; ExternalWritable := 'False'} : Bool;
      Temp_Rückwärts { ExternalAccessible := 'False'; ExternalVisible := 'False'; ExternalWritable := 'False'} : Bool;
      Temp_Bremse { ExternalAccessible := 'False'; ExternalVisible := 'False'; ExternalWritable := 'False'} : Bool;
   END_VAR


BEGIN
	(*
	    Drehtelleransteuerung
	    =========================================
	    created: 23.09.2021 Franz Zwirglmaier 
	    
	    
	  
	*)
	
	
	
	REGION Störungen
	    // Störung Drehteller dreht nicht ********************************
	    #Timer_Drehteller_Laufzeit(IN := #Schuetz_links OR #Schuetz_rechts,
	                               PT := #Time_Drehteller_Laufzeit);
	    
	    IF #Timer_Drehteller_Laufzeit.Q THEN
	        #SM_Drehteller_dreht_nicht := TRUE;
	    ELSE
	        IF #SM_reset THEN
	            #SM_Drehteller_dreht_nicht := FALSE;
	        END_IF;
	    END_IF;
	    //****************************************************************
	    
	    
	    // Störmeldung Drehteller nicht in Position ***********************
	    #Timer_Drehteller_nicht_in_Position(IN := #Schuetz_links = FALSE AND #Schuetz_rechts = FALSE AND #ES_in_Position = FALSE AND #iStep = 10 ,
	                                        PT := #Time_Drehteller_nicht_in_Position);
	    
	    
	    IF #Timer_Drehteller_nicht_in_Position.Q THEN
	        #SM_Drehteller_nicht_in_Position := TRUE;
	    ELSE
	        IF #SM_reset THEN
	            #SM_Drehteller_nicht_in_Position := FALSE;
	        END_IF;
	    END_IF;
	    //****************************************************************
	    
	    
	    // Störmeldung Motorschutz ***************************************
	    IF #Motorschutz = false THEN
	        #SM_Motorschutz := true;
	    ELSE
	        IF #SM_reset THEN
	            #SM_Motorschutz := false;
	        END_IF;
	    END_IF;
	    //****************************************************************
	    
	    // Störmeldung Sicherheitsbit ***************************************
	    IF #Sicherheitsbit_DT= false AND
	        #Befehlsfreigabe THEN
	        #SM_Sicherheitsbit := true;
	    ELSE
	        IF #SM_reset THEN
	            #SM_Sicherheitsbit := false;
	        END_IF;
	    END_IF;
	    //****************************************************************
	    
	    
	    
	    
	    
	END_REGION
	
	
	
	
	
	
	
	REGION Wartungszähler
	    // Aktorenzyklen zählen **************************************************
	    #F_TRIG_Zyklenzähler(CLK := #Schuetz_links OR #Schuetz_rechts);
	    IF #F_TRIG_Zyklenzähler.Q THEN
	        #Aktorzyklen := #Aktorzyklen + 1;
	    END_IF;
	    
	    
	    // Wartungszähler ***************************************
	    #Modolo_Wartungszähler := #Aktorzyklen MOD #Wartungsintervall;
	    #F_TRIG_Modolo_gleich_0(CLK := #Modolo_Wartungszähler = 0);
	    IF #F_TRIG_Modolo_gleich_0.Q THEN
	        #SM_Wartung := true;
	    ELSE
	        IF #SM_reset THEN
	            #SM_Wartung := false;
	        END_IF;
	    END_IF;
	    //****************************************************************
	END_REGION
	
	
	REGION Befehlsfreigabe
	    IF #Automatik AND #Ablauf_aktiv THEN
	        IF #Auto_Frg_Drehen_Vorwärts THEN
	            #Befehlsfreigabe := TRUE;
	        END_IF;
	    END_IF;
	    
	    IF #Manuell AND #Manuellfreigabe THEN
	        IF #Manu_Frg_Drehen_Vorwärts THEN
	            #Befehlsfreigabe := TRUE;
	        END_IF;
	    END_IF;
	    
	    IF #Richten AND #Richtenfreigabe THEN
	        IF #Richt_Frg_Drehen_Vorwärts THEN
	            #Befehlsfreigabe := TRUE;
	        END_IF;
	    END_IF;
	    
	    
	    IF #Automatik = false AND
	        #Manuell = false AND
	        #Richten = false THEN
	        #iStep := 0;
	        #Befehlsfreigabe := FALSE;
	    END_IF;
	    
	    
	    IF #SM_Motorschutz OR
	        #SM_Sicherheitsbit THEN
	        #iStep := 0;
	        #Befehlsfreigabe := FALSE;
	    END_IF;
	    
	    
	    
	END_REGION
	
	
	REGION Automatikablauf
	    
	    // Timer Öffnungszeit Bremse **************************************
	    #Timer_Öffnungszeit_Bremse(IN := #Schrittkette_start,
	                               PT := #Time_Öffnungszeit_Bremse);
	    
	    
	    // Timer Startzeit **************************************
	    #Timer_Startzeit(IN := #Schuetz_rechts OR #Schuetz_links,
	                     PT := #Time_Startzeit);
	    
	    
	    
	    
	    //************************ Automatikschrittkette ******************
	    
	    
	    
	    
	    
	    // *********Initialisieren*****************************************
	    IF #SM_Motorschutz OR
	        #SM_Sicherheitsbit OR
	        #SM_Drehteller_nicht_in_Position OR
	        #SM_Drehteller_dreht_nicht   THEN
	        #iStep := 0;
	        #Temp_Vorwärts := false;
	        #Temp_Rückwärts := false;
	        #Temp_Bremse := false;
	        #Fertigmeldung_Drehteller := false;
	        #Auto_Frg_Drehen_Vorwärts := 0;
	        #Auto_Frg_Drehen_Rückwärts:= 0;
	        
	    END_IF;
	    // *****************************************************************
	    
	    
	    
	    // Schrittkette starten
	    IF #Befehlsfreigabe THEN
	        #Schrittkette_start := true;
	    ELSE
	        #iStep := 0;
	        //#Temp_Bremse := FALSE;
	    END_IF;
	    
	    
	    CASE #iStep OF
	        0:
	            // =========================================================
	            // Schritt 1 : Start, Bremse öffnen
	            // =========================================================
	            IF #Schrittkette_start THEN
	                #iStep := 5;
	                
	              
	            END_IF;
	            
	        5:
	            // =========================================================
	            // Schritt 2 : Drehteller vorwärts oder Rückwärts
	            // =========================================================
	            IF #Timer_Öffnungszeit_Bremse.Q THEN
	                #iStep := 10;
	                #Schrittkette_start := false;
	                #Befehlsfreigabe := false;
	                #Fertigmeldung_Drehteller := false;
	                
	                IF #links0_rechts1_drehen THEN
	                    #Temp_Vorwärts := TRUE;
	                    #Temp_Bremse := TRUE;
	                ELSE
	                    #Temp_Rückwärts := TRUE;
	                    #Temp_Bremse := TRUE;
	                END_IF;
	               
	            END_IF;
	            
	        10:
	            // =========================================================
	            // Schritt 3 :  Position erreicht
	            // =========================================================
	            IF #Timer_Startzeit.Q AND
	                #ES_in_Position THEN
	                #iStep := 15;
	                #Temp_Vorwärts := FALSE;
	                #Temp_Rückwärts := FALSE;
	                #Temp_Bremse := FALSE;
	            END_IF;
	            
	        15:
	            // =========================================================
	            // Schritt 4 :  Fertig
	            // =========================================================
	            IF #ES_in_Position THEN
	                #iStep := 0;
	                
	                #Befehlsfreigabe := false;
	                #Auto_Frg_Drehen_Vorwärts := false;
	                #Auto_Frg_Drehen_Rückwärts := false;
	                #Manu_Frg_Drehen_Vorwärts := false;
	                #Manu_Frg_Drehen_Rückwärts := false;
	                #Richt_Frg_Drehen_Vorwärts := false;
	                #Richt_Frg_Drehen_Rückwärts := false;
	                #Temp_Bremse := false;
	                #Fertigmeldung_Drehteller := true;
	                
	                
	            END_IF;
	            
	    END_CASE;
	    
	END_REGION
	
	REGION Befehlsausgabe
	    #Schuetz_rechts  :=  #Temp_Vorwärts;
	    #Schuetz_links :=  #Temp_Rückwärts;
	    #DT_Bremse:=  #Temp_Bremse;
	END_REGION
	    
	
END_FUNCTION_BLOCK

FUNCTION_BLOCK "Wendelförderer"
{ S7_Optimized_Access := 'TRUE' }
VERSION : 0.1
   VAR_INPUT 
      LS_Teil_vorhanden : Bool;
      LS_Puffer_voll : Bool;
      Pufferzeit : Time;
      Vorlaufzeit_abblasen : Time;
      Nachlaufzeit_abblasen : Time;
      LFZ_Bunker_SM : Time;
      Topf_leer : Bool;
      ACK : Bool;
      LS_Hell_Dunkel_aktiv : Bool;
      LFZ_Puffer_SM : Time;
      VZ_Teil_vorhanden : Time;
      Nachlaufzeit_Bunker : Time;
      Automatik : Bool;
      Manuell : Bool;
      LFZ_Teile_SM : Time;
   END_VAR

   VAR_OUTPUT 
      WF_Start : Bool;
      Linearfoerderer_Start : Bool;
      SM_LS_Teileerkennung : Bool;
      SM_Bunker : Bool;
      Bunker_Start : Bool;
      SM_LS_Puffer : Bool;
   END_VAR

   VAR_IN_OUT 
      WF_abblasen : Bool;
   END_VAR

   VAR 
      TON_WF_HT {InstructionName := 'TON_TIME'; LibVersion := '1.0'} : TON_TIME;
      TON_WF_Freigabe {InstructionName := 'TON_TIME'; LibVersion := '1.0'} : TON_TIME;
      WF_Freigabe : Bool;
      TON_WF_Stop {InstructionName := 'TON_TIME'; LibVersion := '1.0'} : TON_TIME;
      TON_WF_abblasen_Vorlauf {InstructionName := 'TON_TIME'; LibVersion := '1.0'} : TON_TIME;
      Nachlauf_Start : Bool;
      TON_WF_abblasen_Nachlauf {InstructionName := 'TON_TIME'; LibVersion := '1.0'} : TON_TIME;
      TON_Bunker_Aus {InstructionName := 'TON_TIME'; LibVersion := '1.0'} : TON_TIME;
      TON_Topf_leer {InstructionName := 'TON_TIME'; LibVersion := '1.0'} : TON_TIME;
      TON_SM_Puffer {InstructionName := 'TON_TIME'; LibVersion := '1.0'} : TON_TIME;
      TON_LS_Teil_vorhanden {InstructionName := 'TON_TIME'; LibVersion := '1.0'} : TON_TIME;
      LS_Teil_vorhanden_mit_VZ : Bool;
      TON_SM_Teile {InstructionName := 'TON_TIME'; LibVersion := '1.0'} : TON_TIME;
      TON_SM_Bunker {InstructionName := 'TON_TIME'; LibVersion := '1.0'} : TON_TIME;
      Bunker_fertig : Bool;
      HM_LS_Dunkel : Bool;
      F_TRIG_Hell_Dunkel_aktiv {InstructionName := 'F_TRIG'; LibVersion := '1.0'} : F_TRIG;
      SM_LS_Hell_Dunkel : Bool;
      HM_Topf_leer : Bool;
      HM_leer_nach_Zeit : Bool;
      F_TRIG_1 {InstructionName := 'F_TRIG'; LibVersion := '1.0'} : F_TRIG;
      F_TRIG_2 {InstructionName := 'F_TRIG'; LibVersion := '1.0'} : F_TRIG;
   END_VAR


BEGIN
	    (*---------------------------WF Freigabe------------------------*)
	#TON_WF_HT(IN := NOT #LS_Teil_vorhanden,
	           PT := t#5s);
	
	
	#TON_WF_Freigabe(IN := NOT #LS_Puffer_voll OR #TON_WF_HT.Q, PT := T#10ms);
	
	IF (#Automatik OR #Manuell) AND #TON_WF_Freigabe.Q THEN
	    #WF_Freigabe := 1;
	END_IF;
	
	#TON_WF_Stop(IN := #LS_Puffer_voll, PT := #Pufferzeit);
	
	IF #TON_WF_Stop.Q OR NOT (#Automatik OR #Manuell) THEN
	    #WF_Freigabe := 0;
	END_IF;
	
	
	(*---------------------------Teile abblasen---------------------*)
	
	(*Vorlaufzeit*)
	#TON_WF_abblasen_Vorlauf(IN:= #WF_abblasen, PT:=#Vorlaufzeit_abblasen);
	
	(*Nachlaufzeit*)
	
	#F_TRIG_2(CLK:= #WF_Start);
	
	IF #F_TRIG_2.Q THEN
	    #Nachlauf_Start := 1;
	END_IF;
	
	IF #TON_WF_abblasen_Nachlauf.Q THEN
	    #Nachlauf_Start := 0;
	END_IF;
	
	#TON_WF_abblasen_Nachlauf(IN:= #Nachlauf_Start, PT:=#Nachlaufzeit_abblasen);
	
	(*Abblasen*)
	IF #WF_Freigabe THEN
	    #WF_abblasen := 1;
	END_IF;
	
	
	#F_TRIG_1(CLK:= #Nachlauf_Start);
	
	IF #F_TRIG_1.Q THEN
	    #WF_abblasen := 0;
	END_IF;
	
	
	(*---------------------------WF Ein-----------------------------*)
	
	IF  #WF_Freigabe AND NOT #SM_LS_Teileerkennung THEN
	    #WF_Start := 1;
	ELSE
	    #WF_Start := 0;
	END_IF;
	
	
	(*---------------------------Linearförderer---------------------*)
	
	IF (#Manuell OR #Automatik) THEN
	    #Linearfoerderer_Start := 1;
	ELSE
	    #Linearfoerderer_Start := 0;
	END_IF;
	
	(*-----------------------Bunker---------------------------------*)
	IF #Topf_leer AND #WF_Start AND NOT #HM_leer_nach_Zeit AND NOT #SM_Bunker THEN
	    #HM_Topf_leer := 1;
	ELSE
	    #HM_Topf_leer := 0;
	END_IF;
	
	#TON_Topf_leer(IN:=#HM_Topf_leer, PT:=t#5s);
	
	IF #TON_Topf_leer.Q THEN
	    #HM_leer_nach_Zeit := 1;
	END_IF;
	
	IF #TON_Bunker_Aus.Q THEN
	    #HM_leer_nach_Zeit := 0;
	    #Bunker_fertig := 1;
	END_IF;
	
	#TON_Bunker_Aus(IN := #HM_leer_nach_Zeit, PT := #Nachlaufzeit_Bunker);
	
	IF (#Automatik OR #Manuell) AND #HM_leer_nach_Zeit THEN
	    #Bunker_Start := 1;
	ELSE
	    #Bunker_Start := 0;
	END_IF;
	
	(*-----------------------Störungen------------------------------*)
	
	
	(*Laufzeitüberwachung LS Teileerkennung*)
	#TON_SM_Teile(IN := (#WF_Start OR #LS_Puffer_voll) AND NOT #LS_Teil_vorhanden AND NOT #SM_LS_Teileerkennung, PT := #LFZ_Teile_SM);
	
	IF #TON_SM_Teile.Q THEN
	    #SM_LS_Teileerkennung := TRUE;
	END_IF;
	
	IF #SM_LS_Teileerkennung AND #ACK THEN
	    #SM_LS_Teileerkennung := FALSE;
	END_IF;
	
	(*Laufzeitüberwachung Bunker*)
	#TON_SM_Bunker(IN := (#Bunker_fertig AND #WF_Start AND #Topf_leer), PT := #LFZ_Bunker_SM);
	
	IF #Bunker_fertig AND #WF_Start AND NOT #Topf_leer THEN
	    #Bunker_fertig := FALSE;
	END_IF;
	
	IF #TON_SM_Bunker.Q THEN
	    #SM_Bunker := TRUE;
	END_IF;
	
	IF #SM_Bunker AND #ACK THEN
	    #SM_Bunker := FALSE;
	    #Bunker_fertig := TRUE;
	END_IF;
	
	(*Laufzeitüberwachung LS PUFFER*)
	#TON_SM_Puffer(IN := #WF_Start AND NOT #Topf_leer AND NOT #ACK, PT := #LFZ_Puffer_SM);
	
	IF #TON_SM_Puffer.Q THEN
	    #SM_LS_Puffer := TRUE;
	END_IF;
	
	IF #SM_LS_Puffer AND #ACK THEN
	    #SM_LS_Puffer := FALSE;
	END_IF;
	
	(*VZ_LS_Teilvorhanden*)
	
	#TON_LS_Teil_vorhanden(IN:= #LS_Teil_vorhanden AND NOT #SM_LS_Hell_Dunkel, PT:= #VZ_Teil_vorhanden);
	
	IF #TON_LS_Teil_vorhanden.Q THEN
	    #LS_Teil_vorhanden_mit_VZ := TRUE;
	ELSE
	    #LS_Teil_vorhanden_mit_VZ := FALSE;
	END_IF;
	
	(*SM_Lichtschranke nicht Hell_Dunkel geworden*)
	(*Wird ausgelöst wenn die Aktivierung null wird und die Lichtschranke nicht null war*)
	IF (#LS_Hell_Dunkel_aktiv AND NOT #LS_Teil_vorhanden) THEN
	    #HM_LS_Dunkel := TRUE;
	END_IF;
	
	#F_TRIG_Hell_Dunkel_aktiv(CLK:= #LS_Hell_Dunkel_aktiv);
	
	IF (#F_TRIG_Hell_Dunkel_aktiv.Q AND NOT #HM_LS_Dunkel) THEN
	    #SM_LS_Hell_Dunkel := TRUE;
	END_IF;
	
	IF (NOT #LS_Hell_Dunkel_aktiv AND #SM_LS_Hell_Dunkel AND #ACK) THEN
	    #SM_LS_Hell_Dunkel := FALSE;
	END_IF;
END_FUNCTION_BLOCK

FUNCTION "2CharToUInt" : Void
{ S7_Optimized_Access := 'TRUE' }
VERSION : 0.1
   VAR_INPUT 
      Zehner : Char;
      Einer : Char;
   END_VAR

   VAR_OUTPUT 
      OUT_Int : Int;
   END_VAR

   VAR_TEMP 
      tempZ : Char;
      Result : UInt;
   END_VAR


BEGIN
	IF #Zehner = ' ' OR #Zehner = Char#0 THEN
	    #tempZ := '0';
	ELSE
	    #tempZ := #Zehner;
	END_IF;
	
	IF #tempZ < '0' OR #tempZ > '9' OR #Einer < '0' OR #Einer > '9' THEN
	    #Result := 0;
	ELSE
	    #Result := (CHAR_TO_UINT(#tempZ) - CHAR_TO_UINT('0')) * 10 + CHAR_TO_UINT(#Einer) - CHAR_TO_UINT('0');
	END_IF;
	#OUT_Int := UINT_TO_INT( #Result);
	
	
END_FUNCTION

FUNCTION_BLOCK "Messtechnik Arbeitsstellungserkennung"
{ S7_Optimized_Access := 'TRUE' }
VERSION : 0.1
   VAR_INPUT 
      Messwert : Real;
      Start : Bool;
      Startverzögerung_Time : Time;
      Auswerteintervalle : Int;
      Auswertetoleranz : Real;
   END_VAR

   VAR_OUTPUT 
      AS_Erreicht : Bool;
   END_VAR

   VAR 
      TON_1 {InstructionName := 'TON_TIME'; LibVersion := '1.0'; S7_SetPoint := 'False'} : TON_TIME;
      TON_2 {InstructionName := 'TON_TIME'; LibVersion := '1.0'; S7_SetPoint := 'False'} : TON_TIME;
      R_TRIG {InstructionName := 'R_TRIG'; LibVersion := '1.0'; S7_SetPoint := 'False'} : R_TRIG;
      Startverzögerung {InstructionName := 'TON_TIME'; LibVersion := '1.0'; S7_SetPoint := 'False'} : TON_TIME;
      x_Wert : Array[0..200] of Real;
      i : Int;
      Static_Auswerteintervalle : Int;
   END_VAR


BEGIN
	(/*
	    Messtechnik Arbeitsstellungserkennung
	    =========================================
	    created: 27.05.2022 Franz Zwirglmaier 
	
	
	 Beschreibung:
	 Mit dem Start-Eingang wird Messwert in einer Abtastfrequenz von 100Hz aufgezeichnet.
	 Nach der in der "Startverzögerung_Time" eingestellten Zeit werden die Anzahl der Aufgezeichneten Werte,
	 die im Parameter "Auswerteintervalle" eingestellt sind, ausgewertet.
	 Liegen die ausgewerteten Werte innerhalb der vorgegebenen Auswertetoleranz, wird der Ausgang "AS_Erreicht" gesetzt.  
	
	
	*/)
	
	
	
	// Abtastfrequenz 100Hz = 10ms 
	#TON_1(IN := NOT #TON_2.Q,
	           PT := T#5ms);
	    #TON_2(IN := #TON_1.Q,
	           PT := T#5ms);
	#R_TRIG(CLK := #TON_1.Q);
	    
	    
	// Startverzögerung 
	#Startverzögerung(IN := #Start, PT := #Startverzögerung_Time);
	
	IF #Start THEN
	// Messwert aufzeichnen    
	    #x_Wert[0] := #Messwert;
	    
	    IF #R_TRIG.Q THEN
	        FOR #i := 0 TO 99 DO
	            #x_Wert[100-#i] := #x_Wert[99-#i];
	        END_FOR;
	    END_IF;
	    
	    
	// Auswerteintervalle Begrenzen
	    IF #Auswerteintervalle > 100 THEN
	        #Static_Auswerteintervalle := 100;
	    ELSE
	        #Static_Auswerteintervalle := #Auswerteintervalle;
	    END_IF;
	    
	// Auswertung   
	    FOR #i := 1 TO #Static_Auswerteintervalle DO
	        IF #Startverzögerung.Q AND (ABS_REAL(#x_Wert[0] - #x_Wert[#i]) < #Auswertetoleranz) THEN
	            #AS_Erreicht := true;
	        ELSE
	            #AS_Erreicht := false;
	            EXIT;
	        END_IF;
	    END_FOR;
	ELSE
	    FOR #i := 0 TO 100 DO
	        #x_Wert[#i] := 0.0;
	    END_FOR;
	    #AS_Erreicht := false;
	    #TON_1.IN := false;
	    #TON_2.IN := false;
	END_IF;
	
	
	        
	            
END_FUNCTION_BLOCK

FUNCTION "Stringcopy" : Void
{ S7_Optimized_Access := 'TRUE' }
VERSION : 0.1
   VAR_INPUT 
      InString : WString;
   END_VAR

   VAR_OUTPUT 
      OutString : WString;
   END_VAR


BEGIN
	
	//
	// String umkopieren
	//
	
	// Anweisungsteil
	#OutString := #InString;
	
	
END_FUNCTION

FUNCTION_BLOCK "Taktzeitermittlung_Start_V1_0"
TITLE = Taktzeitermittlung_Start
{ S7_Optimized_Access := 'TRUE' }
AUTHOR : FA
VERSION : 1.0
//Ausgabe der Zeit zwischen 2 Starttriggern 27.03.2024 FA
   VAR_INPUT 
      E_Starttrigger : Bool;
   END_VAR

   VAR_OUTPUT 
      A_letzteZykluszeit : Time;
   END_VAR
   VAR_OUTPUT DB_SPECIFIC
      A_letze10Zyklen : Array[0..10] of Time := [T#1MS, T#765MS, T#759MS, T#762MS, T#758MS, T#763MS, T#768MS, T#763MS, T#766MS, T#757MS, T#766MS];
   END_VAR

   VAR 
      Flanke_Takt {InstructionName := 'R_TRIG'; LibVersion := '1.0'} : R_TRIG;
      aktuelle_Zeit { S7_SetPoint := 'True'} : LDT;
      letzte_Zeit : LDT;
      Read_Time : Int;
      Taktzeit : Time;
      Zykluszeit_temp : Time;
      "10_Zyklen" : Array[0..10] of Time;
   END_VAR

   VAR_TEMP 
      i : Int;
   END_VAR


BEGIN
	
	(*
	Zeit zwischen Flanke am Triggereingang zum nächsten Flanke wird ermittelt und am Ausgang letzte Zykluszeit ausgegeben
	zusätzlichwerden die letzten 10 Zykluszeiten am Ausgangangsarray ausgegeben *)
	
	REGION Taktzeit
	    
	    #Flanke_Takt(CLK := #E_Starttrigger);
	    IF #Flanke_Takt.Q THEN
	        #Zykluszeit_temp := t#0s;
	        #letzte_Zeit := #aktuelle_Zeit;
	        #Read_Time := RD_SYS_T(#aktuelle_Zeit);
	        #Taktzeit := LTIME_TO_TIME(LDT_TO_LTIME(T_SUB(IN1 := #aktuelle_Zeit, IN2 := #letzte_Zeit)));
	        #"10_Zyklen"[0] := #Taktzeit;
	        FOR #i := 10 TO 1 BY - 1 DO
	            #"10_Zyklen"[#i] := #"10_Zyklen"[#i - 1]
	            ;
	        END_FOR;
	        
	        #A_letzteZykluszeit :=  #"10_Zyklen"[1];
	        #A_letze10Zyklen := #"10_Zyklen";
	    END_IF;
	END_REGION
END_FUNCTION_BLOCK

FUNCTION "GIT_TEstbaustein" : Void
{ S7_Optimized_Access := 'TRUE' }
VERSION : 0.1
   VAR_INPUT 
      IN_1 : Bool;
      IN_2 : Bool;
   END_VAR

   VAR_OUTPUT 
      OUT_1 : Bool;
   END_VAR


BEGIN
	IF #IN_1 THEN
	    #OUT_1 := true;
	END_IF;
	
	
	IF #IN_2 THEN
	    #OUT_1 := true;
	END_IF;
	
	
END_FUNCTION

FUNCTION "GIT_Testbaustein 2" : Void
{ S7_Optimized_Access := 'TRUE' }
VERSION : 0.1
   VAR_INPUT 
      Input_REAL1 : Real;
      Input_REAL2 : Real;
   END_VAR

   VAR_OUTPUT 
      Ouput_REAL1 : Real;
      Ouput_REAL2 : Real;
   END_VAR

   VAR_TEMP 
      Bool1 : Bool;
   END_VAR


BEGIN
	REGION Testregion
	    // Statement section REGION
	    // 
	    IF #Bool1 THEN
	        #Ouput_REAL2 := #Input_REAL1 + #Input_REAL2;
	        
	    END_IF;
	    
	    
	END_REGION
	
	
	REGION Testregion2
	    // Statement section REGION
	    // 
	    IF #Bool1 THEN
	        #Ouput_REAL1 := #Input_REAL1 - #Input_REAL2;
	        
	    END_IF;
	    
	    
	END_REGION
END_FUNCTION

DATA_BLOCK "DB002_LabView_DB"   // DB3
// stored: InstanceOfName FB002_LabView, InstanceOfType FB
"FB002_LabView"
BEGIN
END_DATA_BLOCK

DATA_BLOCK "DataFromSafey_DB"   // DB70
// stored: AssignedProDiagFB ProDiag_Allgemein, InstanceOfName DataFromSafey, InstanceOfType FB
"DataFromSafey"
BEGIN
END_DATA_BLOCK

DATA_BLOCK "DataToSafety_DB"   // DB52
// stored: InstanceOfName DataToSafety, InstanceOfType FB
"DataToSafety"
BEGIN
END_DATA_BLOCK

DATA_BLOCK "Main_Safety_RTG1_DB"   // DB15, F_DB
NAME : FUSI
// stored: InstanceOfName Main_Safety_RTG1, InstanceOfType FB
"Main_Safety_RTG1"
BEGIN
END_DATA_BLOCK

DATA_BLOCK "Zaehler_Sicherheit_DB"   // DB203
// stored: InstanceOfName Zaehler_Sicherheit, InstanceOfType FB
"Zaehler_Sicherheit"
BEGIN
END_DATA_BLOCK

DATA_BLOCK "02_Wartungsfreigaben_DB"   // DB22
// stored: InstanceOfName 02_Wartungsfreigaben, InstanceOfType FB
"02_Wartungsfreigaben"
BEGIN
END_DATA_BLOCK

DATA_BLOCK "03_Betriebsart_DB"   // DB11
// stored: InstanceOfName 03_Betriebsart, InstanceOfType FB
"03_Betriebsart"
BEGIN
END_DATA_BLOCK

DATA_BLOCK "05_Not-Aus_DB"   // DB164
// stored: InstanceOfName 05_Not-Aus, InstanceOfType FB
"05_Not-Aus"
BEGIN
END_DATA_BLOCK

DATA_BLOCK "06_Grundstellungen_DB"   // DB177
// stored: InstanceOfName 06_Grundstellungen, InstanceOfType FB
"06_Grundstellungen"
BEGIN
END_DATA_BLOCK

DATA_BLOCK "08_Systemzeit_DB"   // DB29
// stored: InstanceOfName 08_Systemzeit, InstanceOfType FB
"08_Systemzeit"
BEGIN
END_DATA_BLOCK

DATA_BLOCK "Leuchtmelder Ampel_DB"   // DB77
// stored: InstanceOfName Leuchtmelder Ampel, InstanceOfType FB
"Leuchtmelder Ampel"
BEGIN
   Ampelbaustein_MG_Instance.Sammelstoerung := FALSE;
   Ampelbaustein_MG_Instance.BA_0 := FALSE;
   Ampelbaustein_MG_Instance.BA_A := FALSE;
   Ampelbaustein_MG_Instance.BA_M := TRUE;
   Ampelbaustein_MG_Instance.BA_R := FALSE;
   Ampelbaustein_MG_Instance.BA_V := FALSE;
   Ampelbaustein_MG_Instance.Ablauf_ist_aktiv := FALSE;
   Ampelbaustein_MG_Instance.Blinker := FALSE;
   Ampelbaustein_MG_Instance.Ampel_rot := FALSE;
   Ampelbaustein_MG_Instance.Ampel_gelb := FALSE;
   Ampelbaustein_MG_Instance.Ampel_gruen := FALSE;
   Ampelbaustein_MG_Instance.Akkustik := FALSE;
   Ampelbaustein_MG_Instance.Timer_Hupe_EIN.PT := T#5M;
   Ampelbaustein_MG_Instance.Timer_Hupe_EIN.IN := FALSE;
   Ampelbaustein_MG_Instance.Timer_Hupe_Aus.PT := T#10M;
   Ampelbaustein_MG_Instance.Timer_Hupe_Aus.IN := FALSE;
   Ampelbaustein_MG_Instance.Ampel_Zustand := 0;
END_DATA_BLOCK

DATA_BLOCK "Melden_VisuAllgemein_DB"   // DB155
// stored: InstanceOfName Melden_VisuAllgemein, InstanceOfType FB
"Melden_VisuAllgemein"
BEGIN
END_DATA_BLOCK

DATA_BLOCK "01_Alle_Zaehler_DB"   // DB162
// stored: AssignedProDiagFB Pos12_ProDiag, InstanceOfName 01_Alle_Zaehler, InstanceOfType FB
"01_Alle_Zaehler"
BEGIN
END_DATA_BLOCK

DATA_BLOCK "02_Wartungszaehler_DB"   // DB4
AUTHOR : Falter
FAMILY : HMI
VERSION : 1.0
// stored: InstanceOfName 02_Wartungszaehler, InstanceOfType FB
"02_Wartungszaehler"
BEGIN
END_DATA_BLOCK

DATA_BLOCK "Verwaltung_Teiledaten_FB_DB"   // DB1
// stored: InstanceOfName Verwaltung_Teiledaten_FB, InstanceOfType FB
"Verwaltung_Teiledaten_FB"
BEGIN
END_DATA_BLOCK

DATA_BLOCK "POS3_0_Antriebe_DB"   // DB24
// stored: AssignedProDiagFB POS3_0_Prodiag, InstanceOfName POS3_0_Antriebe, InstanceOfType FB
"POS3_0_Antriebe"
BEGIN
END_DATA_BLOCK

DATA_BLOCK "POS3_0_Melden_Visu_DB"   // DB62
// stored: AssignedProDiagFB POS3_0_Prodiag, InstanceOfName POS3_0_Melden_Visu, InstanceOfType FB
"POS3_0_Melden_Visu"
BEGIN
END_DATA_BLOCK

DATA_BLOCK "POS3_0_Messtechnik_DB"   // DB60
// stored: AssignedProDiagFB POS4_0_Prodiag, InstanceOfName POS3_0_Messtechnik, InstanceOfType FB
"POS3_0_Messtechnik"
BEGIN
END_DATA_BLOCK

DATA_BLOCK "POS3_0_SK_Ablauf_DB"   // DB35
// stored: AssignedProDiagFB POS3_0_Prodiag, InstanceOfName POS3_0_SK_Ablauf, InstanceOfType FB
"POS3_0_SK_Ablauf"
BEGIN
END_DATA_BLOCK
